{region 'Documentation'}
(*!
<summary>Calls Preparations and supplies their scenario-specific combined observations.</summary>
<description>
Called after ProcessAbort on every initialized call except Completed, with the current
Preparation-phase Enable. Call Preparations even when disabled so their observations and
deactivation remain correct; report the combination through UpdatePreparationStatus.

Only enabled phase processing may advance through NextPreparationState or
CompletePreparations. After entry into Test states, loss of Preparation Ready or Completed is not by
itself a Test Case failure. This abstract hook has no base implementation.
</description>
*)
{endregion}
METHOD PROTECTED ABSTRACT ProcessPreparations
VAR_INPUT
    Enable: BOOL; //! TRUE while this hook's lifecycle phase is active; FALSE must not advance that phase.
END_VAR
(* Example: declare a local ObservedStatus : ST_PreparationStatus; combine multiple Preparations as needed.
MyPreparation(Enable := Enable);
ObservedStatus := MyPreparation.Status;
UpdatePreparationStatus(Ready := ObservedStatus.Ready,
    Running := ObservedStatus.Running,
    Completed := ObservedStatus.Completed,
    HasError := ObservedStatus.Error,
    State := ObservedStatus.State);
IF Enable AND FPreparationStatus.Completed AND NOT FPreparationStatus.Error THEN
    CompletePreparations();
END_IF;
*)
END_METHOD

{region 'Documentation'}
(*!
<summary>Consumes same-task requests, reports each received request and prioritizes Reset &gt; Abort &gt; Start.</summary>
<description>
Discards requests before initialization; never changes lifecycle state.
</description>
*)
{endregion}
METHOD PRIVATE ProcessRequests
VAR_IN_OUT
    InputRequests : ST_Command; //! Same-task request mailbox consumed and cleared, including calls made before successful initialization.
END_VAR
VAR_OUTPUT
    Requests : ST_Command; //! Qualified request snapshot with Reset over Abort over Start; all FALSE before initialization.
END_VAR
Requests.Reset := FALSE;
Requests.Abort := FALSE;
Requests.Start := FALSE;

IF NOT FInitialized THEN
    InputRequests.Reset := FALSE;
    InputRequests.Abort := FALSE;
    InputRequests.Start := FALSE;
    RETURN;
END_IF;

Requests.Reset := InputRequests.Reset;
Requests.Abort := InputRequests.Abort AND NOT InputRequests.Reset;
Requests.Start := InputRequests.Start AND NOT InputRequests.Abort AND NOT InputRequests.Reset;

IF InputRequests.Reset THEN
    PublishEvent(Event := CreateResetEvent(OwnerScope := E_OwnerScope.TestCase,
        Name := FName,
        ResourceName := FResourceName,
        State := FState));
END_IF;

IF InputRequests.Abort THEN
    PublishEvent(Event := CreateAbortEvent(OwnerScope := E_OwnerScope.TestCase,
        Name := FName,
        ResourceName := FResourceName,
        State := FState));
END_IF;

IF InputRequests.Start THEN
    PublishEvent(Event := CreateStartEvent(OwnerScope := E_OwnerScope.TestCase,
        Name := FName,
        ResourceName := FResourceName,
        State := FState));
END_IF;

InputRequests.Reset := FALSE;
InputRequests.Abort := FALSE;
InputRequests.Start := FALSE;
END_METHOD

{region 'Documentation'}
(*!
<summary>Resets owned scenario resources and Assertions during the Reset phase.</summary>
<description>
Called after the base restores the Preparation snapshot to Unknown. Request Assertion resets;
their next regular calls process those requests with bound inputs. Finish through CompleteReset only
once the owned reset work is complete.

Preserve configuration and publisher bindings. One-shot resource protocols must not be
retriggered every cycle. The base owns ResetTimeout; this abstract hook has no base
implementation.
</description>
*)
{endregion}
METHOD PROTECTED ABSTRACT ProcessReset
(* Example: request child resets and observe completion without blocking.
MyAssertion.Reset();
IF OwnedResourcesReset THEN
    CompleteReset();
END_IF;
Issue one-shot resource requests only once if their protocol requires it.
*)
END_METHOD

{region 'Documentation'}
(*!
<summary>Performs scenario actions in the current Test state.</summary>
<description>
Called after ProcessPreparations on every initialized call except Completed. Enable reflects
the phase at invocation, including transitions made by earlier hooks. Keep required cyclic resource
calls active while disabled, but do not advance the Test phase.

Use NextTestState and CompleteTests for immediate transitions. Check errors before successful
completion; do not rely on a previously cached phase flag after changing state. This abstract hook
has no base implementation.
</description>
*)
{endregion}
METHOD PROTECTED ABSTRACT ProcessTests
VAR_INPUT
    Enable: BOOL; //! TRUE while this hook's lifecycle phase is active; FALSE must not advance that phase.
END_VAR
(* Example: keep required cyclic object calls outside the Enable guard.
MyTestObject();
IF NOT Enable THEN
    RETURN;
END_IF;
Perform the action for the current State; check errors before completion.
IF TestCompleted THEN
    CompleteTests();
END_IF;
*)
END_METHOD

{region 'Documentation'}
(*!
<summary>Publishes through the selected instance publisher; the buffer owns lost-event accounting.</summary>
*)
{endregion}
METHOD PRIVATE PublishEvent
VAR_INPUT
    Event : ST_Event; //! Payload copied once through the selected usable publisher, which assigns sequence/time and accounts for loss.
END_VAR
EventPublisher.PublishEvent(Event := Event);
END_METHOD

{region 'Documentation'}
(*!
<summary>Records an Abort request for the next regular FB call.</summary>
<description>
Repeated positive calls coalesce in the same-task request storage. Processing consumes the
requests with priority Reset, Abort, Start; calls before successful initialization are discarded
when processed.

Abort requests controlled termination of execution, not Reset cancellation. The owner
lifecycle determines whether the request applies.
</description>
*)
{endregion}
METHOD PUBLIC RequestAbort
FMethodRequests.Abort := TRUE;
END_METHOD

{region 'Documentation'}
(*!
<summary>Records a Reset request for the next regular FB call.</summary>
<description>
Repeated positive calls coalesce in the same-task request storage. Processing consumes the
requests with priority Reset, Abort, Start; calls before successful initialization are discarded
when processed.

Lifecycle Reset preserves configuration and publisher binding. It is not reinitialization or
Event Buffer Reset; capacity admission belongs to the parent when this object is a child.
</description>
*)
{endregion}
METHOD PUBLIC RequestReset
FMethodRequests.Reset := TRUE;
END_METHOD

{region 'Documentation'}
(*!
<summary>Records a Start request for the next regular FB call.</summary>
<description>
Repeated positive calls coalesce in the same-task request storage. Processing consumes the
requests with priority Reset, Abort, Start; calls before successful initialization are discarded
when processed.

Start is accepted by the lifecycle only in ready Idle. Recording the request does not start
execution synchronously.
</description>
*)
{endregion}
METHOD PUBLIC RequestStart
FMethodRequests.Start := TRUE;
END_METHOD

{region 'Documentation'}
(*!
<summary>Own contribution to the global Event Buffer reservation; changed only with that
aggregate.</summary>
*)
{endregion}
{attribute 'monitoring' := 'call'}
PROPERTY PUBLIC ReservedEntryCount : UINT //! Own contribution to the global Event Buffer reservation; changed only with that aggregate.
GET // PUBLIC
ReservedEntryCount := FReservedEntryCount;
END_GET
END_PROPERTY

{region 'Documentation'}
(*!
<summary>Adjusts this owner's reservation to its execution budget immediately.</summary>
<description>
The budget uses configured state counts and the collected AssertionCountTotal, which must be
valid and stable before Start. Local contribution and publisher accounting are updated together
without a lifecycle transition.

Accepted permits dispatch; WaitingForCapacity is retryable under the owner's timeout; Error
denotes invalid setup or an impossible budget. Calling before initialization reports a Framework
error. Repeated success aligns the total rather than adding a second budget.
</description>
*)
{endregion}
METHOD PUBLIC FINAL ReserveExecutionEvents : E_EventReservationResult //! Accepted on success, WaitingForCapacity for retryable pressure, Error for invalid setup or an impossible budget.
VAR
    EntryCount : UDINT;
END_VAR
VAR CONSTANT
    FixedEventCount : UDINT := 9;
    MaxReservationEntryCount : UDINT := 65535;
END_VAR
ReserveExecutionEvents := E_EventReservationResult.Error;
IF NOT FInitialized THEN
    PublishEvent(Event := CreateFrameworkEvent(Name := FName,
        ResourceName := FResourceName,
        State := FState,
        Severity := E_EventSeverity.Error,
        Message := 'ReserveExecutionEvents requires an initialized Test Case.'));
    RETURN;
END_IF;

EntryCount := INT_TO_UDINT(FPreparationStateCount)
    + INT_TO_UDINT(FTestStateCount)
    + UINT_TO_UDINT(FStatus.AssertionCountTotal)
    + FixedEventCount;
IF EntryCount > MaxReservationEntryCount THEN
    PublishEvent(Event := CreateFrameworkEvent(Name := FName,
        ResourceName := FResourceName,
        State := FState,
        Severity := E_EventSeverity.Error,
        Message := 'Test Case event budget exceeds the reservation range.'));
    RETURN;
END_IF;

ReserveExecutionEvents := UpdateEventReservation(EntryCount := UDINT_TO_UINT(EntryCount),
    HeadroomEntryCount := Param_EventBuffer.EventBufferExecutionHeadroom,
    ConcurrentEntryCount := GVL_Constants.TestSuiteExecutionEventCount);
END_METHOD

{region 'Documentation'}
(*!
<summary>Adjusts this owner's reservation for capacity-admitted Reset immediately.</summary>
<description>
Does not dispatch Reset or clear existing events. Shared headroom and the Suite allowance
participate in admission, not this owner's stored contribution.

Accepted, WaitingForCapacity and Error distinguish success, temporary pressure and invalid
setup. An uninitialized call reports a Framework error. Lifecycle Reset must not silently clear the
reservation.
</description>
*)
{endregion}
METHOD PUBLIC FINAL ReserveResetEvents : E_EventReservationResult //! Accepted on success, WaitingForCapacity for retryable pressure, Error for invalid setup or an impossible budget.
ReserveResetEvents := E_EventReservationResult.Error;
IF NOT FInitialized THEN
    PublishEvent(Event := CreateFrameworkEvent(Name := FName,
        ResourceName := FResourceName,
        State := FState,
        Severity := E_EventSeverity.Error,
        Message := 'ReserveResetEvents requires an initialized Test Case.'));
    RETURN;
END_IF;

ReserveResetEvents := UpdateEventReservation(EntryCount := GVL_Constants.TestCaseResetEventCount,
    HeadroomEntryCount := Param_EventBuffer.EventBufferResetHeadroom,
    ConcurrentEntryCount := GVL_Constants.TestSuiteResetEventCount);
END_METHOD

{region 'Documentation'}
(*!
<summary>Current held Test Case result.</summary>
*)
{endregion}
{attribute 'monitoring' := 'call'}
PROPERTY PUBLIC Result : E_Result //! Current held Test Case result.
GET // PUBLIC
Result := FResult;
END_GET
END_PROPERTY

{region 'Documentation'}
(*!
<summary>Selects lifecycle transitions from requests, observations and timeout supervision.</summary>
*)
{endregion}
METHOD PRIVATE Sequencer
VAR_INPUT
    Requests : ST_Command; //! Consumed request snapshot whose applicability is evaluated against current lifecycle state and error/timeout priority.
END_VAR
VAR
    Message : STRING(GVL_Constants.MessageLength);
END_VAR
IF NOT FInitialized THEN
    IF FState <> E_State.Uninitialized THEN
        ChangeState(NewState := E_State.Uninitialized);
    END_IF;
    RETURN;
END_IF;
IF Requests.Reset THEN
    ChangeState(NewState := E_State.Reset);
END_IF;

CASE FState OF
    E_State.Uninitialized:
        RETURN;

    E_State.Reset:
        IF NOT FStateTimer.IsValid THEN
            PublishEvent(Event := CreateFrameworkEvent(Name := FName,
                ResourceName := FResourceName,
                State := FState,
                Severity := E_EventSeverity.Error,
                Message := 'Task clock error during Test Case reset.'));
            FResult := E_Result.Error;
            ChangeState(NewState := E_State.Completing);
            RETURN;
        END_IF;
        IF FStateTimer.ElapsedLTime >= TIME_TO_LTIME(FConfig.ResetTimeout) THEN
            FHasResetTimeout := TRUE;
            PublishEvent(Event := CreateFrameworkEvent(Name := FName,
                ResourceName := FResourceName,
                State := FState,
                Severity := E_EventSeverity.Error,
                Message := 'Test Case reset timeout reached.'));
            FResult := E_Result.Error;
            ChangeState(NewState := E_State.Completing);
            RETURN;
        END_IF;
        RETURN;

    E_State.Idle:
        IF Requests.Start AND NOT Requests.Abort AND IsReady THEN
            ChangeState(NewState := E_State.Starting);
        END_IF;
        RETURN;

    E_State.Starting:
        IF FResult = E_Result.Error THEN
            ChangeState(NewState := E_State.AbortingFromError);
            RETURN;
        END_IF;
        IF FPreparationStatus.Error THEN
            Message := CONCAT('Preparation error. Preparation state = ', INT_TO_STRING(FPreparationStatus.State));
            Error(Message := Message);
            RETURN;
        END_IF;
        IF FAggregator.Result = E_Result.Error THEN
            Error(Message := 'Test Case evaluation reported Error.');
            RETURN;
        END_IF;
        IF NOT FExecutionTimer.IsValid OR NOT FStateTimer.IsValid THEN
            Error(Message := 'Task clock error.');
            RETURN;
        END_IF;
        IF FExecutionTimer.ElapsedLTime >= TIME_TO_LTIME(FConfig.Timeout) THEN
            FHasTimeout := TRUE;
            Error(Message := 'Test Case timeout.');
            RETURN;
        END_IF;
        IF Requests.Abort THEN
            ChangeState(NewState := E_State.Aborting);
            RETURN;
        END_IF;
        IF (FPreparationStateCount = 0) OR FPreparationStatus.Completed THEN
            ChangeState(NewState := E_State.Running);
            RETURN;
        END_IF;
        ChangeState(NewState := E_State.Preparing);
        RETURN;

    E_State.Preparing..(E_State.Running - 1):
        IF FResult = E_Result.Error THEN
            ChangeState(NewState := E_State.AbortingFromError);
            RETURN;
        END_IF;
        IF NOT IsPreparationActive THEN
            Message := CONCAT('Invalid preparation state = ', INT_TO_STRING(FState));
            Error(Message := Message);
            RETURN;
        END_IF;
        IF FPreparationStatus.Error THEN
            Message := CONCAT('Preparation error. Preparation state = ', INT_TO_STRING(FPreparationStatus.State));
            Error(Message := Message);
            RETURN;
        END_IF;
        IF FAggregator.Result = E_Result.Error THEN
            Error(Message := 'Test Case evaluation reported Error.');
            RETURN;
        END_IF;
        IF NOT FExecutionTimer.IsValid OR NOT FStateTimer.IsValid THEN
            Error(Message := 'Task clock error.');
            RETURN;
        END_IF;
        IF FStateTimer.ElapsedLTime >= TIME_TO_LTIME(FConfig.PreparationTimeout) THEN
            FHasPreparationTimeout := TRUE;
            Message := CONCAT('Preparation timeout. Preparation state = ', INT_TO_STRING(FPreparationStatus.State));
            Error(Message := Message);
            RETURN;
        END_IF;
        IF FExecutionTimer.ElapsedLTime >= TIME_TO_LTIME(FConfig.Timeout) THEN
            FHasTimeout := TRUE;
            Error(Message := 'Test Case timeout.');
            RETURN;
        END_IF;
        IF Requests.Abort THEN
            ChangeState(NewState := E_State.Aborting);
            RETURN;
        END_IF;
        IF (FPreparationStateCount = 0) OR FPreparationStatus.Completed THEN
            ChangeState(NewState := E_State.Running);
            RETURN;
        END_IF;
        // Leave to Running by CompletePreparations
        RETURN;

    E_State.Running..(E_State.Completing - 1):
        IF FResult = E_Result.Error THEN
            ChangeState(NewState := E_State.AbortingFromError);
            RETURN;
        END_IF;
        IF NOT IsTestingActive THEN
            Message := CONCAT('Invalid testing state = ', INT_TO_STRING(FState));
            Error(Message := Message);
            RETURN;
        END_IF;
        IF FAggregator.Result = E_Result.Error THEN
            Error(Message := 'Test Case evaluation reported Error.');
            RETURN;
        END_IF;
        IF NOT FExecutionTimer.IsValid THEN
            Error(Message := 'Task clock error.');
            RETURN;
        END_IF;
        IF FExecutionTimer.ElapsedLTime >= TIME_TO_LTIME(FConfig.Timeout) THEN
            FHasTimeout := TRUE;
            Error(Message := 'Test Case timeout.');
            RETURN;
        END_IF;
        IF Requests.Abort THEN
            ChangeState(NewState := E_State.Aborting);
            RETURN;
        END_IF;
        // Leave to Completing by CompleteTests
        RETURN;

    E_State.Completing:
        ChangeState(NewState := E_State.Completed);
        RETURN;

    E_State.Completed:
        // Leave to Reset on ResetRequested.
        RETURN;

    E_State.Aborting, E_State.AbortingFromError:
        IF NOT FStateTimer.IsValid THEN
            PublishEvent(Event := CreateFrameworkEvent(Name := FName,
                ResourceName := FResourceName,
                State := FState,
                Severity := E_EventSeverity.Error,
                Message := 'Task clock error during Test Case abort.'));
            FResult := E_Result.Error;
            ChangeState(NewState := E_State.Completing);
            RETURN;
        END_IF;
        IF FStateTimer.ElapsedLTime >= TIME_TO_LTIME(FConfig.AbortTimeout) THEN
            FHasAbortTimeout := TRUE;
            PublishEvent(Event := CreateFrameworkEvent(Name := FName,
                ResourceName := FResourceName,
                State := FState,
                Severity := E_EventSeverity.Error,
                Message := 'Test Case abort timeout reached.'));
            FResult := E_Result.Error;
            ChangeState(NewState := E_State.Completing);
            RETURN;
        END_IF;
        IF (FState = E_State.Aborting) AND (FResult = E_Result.Error) THEN
            ChangeState(NewState := E_State.AbortingFromError);
        END_IF;
        RETURN;

    E_State.Aborted, E_State.Error:
        Error(Message := 'Unexpected legacy lifecycle state.');
        RETURN;
ELSE
    Error(Message := 'Unhandled Test Case lifecycle state.');
END_CASE;
END_METHOD

{region 'Documentation'}
(*!
<summary>Current Test Case lifecycle state.</summary>
*)
{endregion}
{attribute 'monitoring' := 'call'}
PROPERTY PUBLIC State : E_State //! Current Test Case lifecycle state.
GET // PUBLIC
State := FState;
END_GET
END_PROPERTY

{region 'Documentation'}
(*!
<summary>Returns the latest Test Case status snapshot without executing children.</summary>
<description>
The base refreshes this snapshot on every FB call, including Uninitialized and Completed.
Assertion counters come from the current collection; the completed owner result remains held.
Runtime is TIME.

Preparation observations are available separately through PreparationStatus. Optional external
publication requires an explicit data wrapper, not access to owner instance data.
</description>
*)
{endregion}
PROPERTY PUBLIC Status : ST_TestCaseStatus //! Returns the latest Test Case status snapshot without executing children.
GET // PUBLIC
Status := FStatus;
END_GET
END_PROPERTY

{region 'Documentation'}
(*!
<summary>Reports the configured maximum number of Test-state entries along one finite lifecycle
path.</summary>
<description>
Set the backing field explicitly in Configure. Before configuration it is
StateCountNotConfigured (-1). Branches use the longest path, including bounded repeated entries;
this is not a count of child instances. Keep it fixed through execution.

At least one Test state is required. CheckInitialization bounds the value by
E_State.Completing - E_State.Running.
</description>
*)
{endregion}
{attribute 'monitoring' := 'call'}
PROPERTY PUBLIC TestStateCount : INT //! Reports the configured maximum number of Test-state entries along one finite lifecycle path.
GET // PUBLIC
TestStateCount := FTestStateCount;
END_GET
END_PROPERTY

{region 'Documentation'}
(*!
<summary>Checks target capacity before changing either reservation count; zero releases without capacity gating.</summary>
<description>
A zero target with no existing contribution succeeds without accessing a publisher. Releasing a nonzero contribution delegates to FreeReservedSpace without a free-capacity check. Positive targets first require valid publisher/accounting and permanent capacity for target plus the concurrent Suite allowance plus headroom. Temporary free capacity uses aggregate minus old own contribution plus target plus headroom; it does not add the Suite allowance again. Even unchanged or reduced positive targets must pass those checks. Failure leaves both ledgers unchanged.
</description>
*)
{endregion}
METHOD PRIVATE UpdateEventReservation : E_EventReservationResult //! Accepted after aligning the own contribution, WaitingForCapacity for temporary pressure, Error for invalid binding/accounting or impossible capacity.
VAR_INPUT
    EntryCount : UINT; //! Target total own reservation, not an additional delta; zero releases the complete own contribution.
    HeadroomEntryCount : UINT; //! Shared unreserved producer headroom included in permanent and temporary capacity checks for a nonzero target.
    ConcurrentEntryCount : UINT; //! Suite allowance used only in the permanent capacity check; actual temporary reservations already include the parent's contribution.
END_VAR
VAR
    Publisher : I_EventPublisher;
    RequiredCapacity : UDINT;
    RequiredFreeEntries : UDINT;
END_VAR
UpdateEventReservation := E_EventReservationResult.Error;
IF (EntryCount = 0) AND (FReservedEntryCount = 0) THEN
    UpdateEventReservation := E_EventReservationResult.Accepted;
    RETURN;
END_IF;

Publisher := EventPublisher;

IF EntryCount = 0 THEN
    IF Publisher.FreeReservedSpace(EntryCount := FReservedEntryCount,
        OwnerReservedEntryCount := FReservedEntryCount) THEN
        UpdateEventReservation := E_EventReservationResult.Accepted;
    END_IF;
    RETURN;
END_IF;

IF NOT Publisher.IsValid THEN
    RETURN;
END_IF;
RequiredCapacity := UINT_TO_UDINT(EntryCount)
    + UINT_TO_UDINT(ConcurrentEntryCount)
    + UINT_TO_UDINT(HeadroomEntryCount);
IF RequiredCapacity > UINT_TO_UDINT(Publisher.Capacity) THEN
    RETURN;
END_IF;
IF FReservedEntryCount > Publisher.ReservedEntryCount THEN
    RETURN;
END_IF;

RequiredFreeEntries := UINT_TO_UDINT(Publisher.ReservedEntryCount)
    - UINT_TO_UDINT(FReservedEntryCount)
    + UINT_TO_UDINT(EntryCount)
    + UINT_TO_UDINT(HeadroomEntryCount);
IF RequiredFreeEntries > UINT_TO_UDINT(Publisher.FreeEntryCount) THEN
    UpdateEventReservation := E_EventReservationResult.WaitingForCapacity;
    RETURN;
END_IF;

IF EntryCount < FReservedEntryCount THEN
    IF Publisher.FreeReservedSpace(EntryCount := FReservedEntryCount - EntryCount,
        OwnerReservedEntryCount := FReservedEntryCount) THEN
        UpdateEventReservation := E_EventReservationResult.Accepted;
    END_IF;
    RETURN;
END_IF;

IF Publisher.ReserveSpace(EntryCount := EntryCount - FReservedEntryCount,
    HeadroomEntryCount := HeadroomEntryCount,
    OwnerReservedEntryCount := FReservedEntryCount) THEN
    UpdateEventReservation := E_EventReservationResult.Accepted;
ELSE
    UpdateEventReservation := E_EventReservationResult.WaitingForCapacity;
END_IF;
END_METHOD

{region 'Documentation'}
(*!
<summary>Replaces the combined Preparation observations without calling children.</summary>
<description>
Combine multiple Preparations according to the concrete scenario; this method imposes no
universal AND/OR aggregation. All supplied flags replace previous observations; Ready is suppressed
while Running.

ExecutionStatus follows Error, Completed, Running, then Idle when Ready and NotReady
otherwise. State is optional diagnostic context, not the owner's phase. Initial/reset Unknown
snapshots are established separately by the base.
</description>
*)
{endregion}
METHOD PROTECTED UpdatePreparationStatus
VAR_INPUT
    Ready : BOOL; //! Resource can be driven to the target state; suppressed while Running. Does not mean target reached.
    Running : BOOL; //! Preparation is actively driving the resource toward its target; forces Ready to FALSE.
    Completed : BOOL; //! Preparation target is currently reached; observation is not latched.
    HasError : BOOL; //! Preparation cannot continue meaningfully; reported as an error observation.
    State : E_State := E_State.Uninitialized; //! Optional combined Preparation state for observation; default Uninitialized.
END_VAR
FPreparationStatus.State := State;
FPreparationStatus.Ready := Ready AND NOT Running;
FPreparationStatus.Running := Running;
FPreparationStatus.Completed := Completed;
FPreparationStatus.Error := HasError;

IF HasError THEN
    FPreparationStatus.ExecutionStatus := E_ExecutionStatus.Error;
ELSIF Completed THEN
    FPreparationStatus.ExecutionStatus := E_ExecutionStatus.Completed;
ELSIF Running THEN
    FPreparationStatus.ExecutionStatus := E_ExecutionStatus.Running;
ELSIF Ready THEN
    FPreparationStatus.ExecutionStatus := E_ExecutionStatus.Idle;
ELSE
    FPreparationStatus.ExecutionStatus := E_ExecutionStatus.NotReady;
END_IF;
END_METHOD

{region 'Documentation'}
(*!
<summary>Applies lifecycle-specific owner result rules to the current aggregate.</summary>
*)
{endregion}
METHOD PRIVATE UpdateResult
IF (FResult = E_Result.Error) AND (FState <> E_State.Uninitialized) THEN
    RETURN;
END_IF;

CASE FState OF
    E_State.Uninitialized, E_State.Starting:
        FResult := E_Result.NotEvaluated;
    E_State.Reset, E_State.Idle:
        RETURN;
    E_State.Aborting:
        IF (FResult = E_Result.Error) OR (FAggregator.Result = E_Result.Error) THEN
            FResult := E_Result.Error;
        ELSE
            FResult := E_Result.Abort;
        END_IF;
    E_State.AbortingFromError:
        FResult := E_Result.Error;
    E_State.Completing:
        IF (FResult = E_Result.Error) OR (FAggregator.Result = E_Result.Error) THEN
            FResult := E_Result.Error;
            RETURN;
        END_IF;
        IF FResult = E_Result.Abort THEN
            RETURN;
        END_IF;
        CASE FAggregator.Result OF
            E_Result.Failed:
                FResult := E_Result.Failed;
            E_Result.Passed, E_Result.NotEvaluated:
                FResult := E_Result.Passed;
        ELSE
            FResult := E_Result.Error;
        END_CASE;
    E_State.Completed:
        RETURN;
ELSE
    IF IsPreparationActive OR IsTestingActive THEN
        FResult := E_Result.NotEvaluated;
    ELSE
        FResult := E_Result.Error;
    END_IF;
END_CASE;
END_METHOD

{region 'Documentation'}
(*!
<summary>Refreshes the typed snapshot from current lifecycle state; does not invoke children.</summary>
*)
{endregion}
METHOD PRIVATE UpdateStatus
VAR
    ExecutionStatus : ST_TestCaseExecutionStatus;
END_VAR
ExecutionStatus.State := FState;
ExecutionStatus.Result := FResult;
ExecutionStatus.ConfigError := FConfigError;
CASE FState OF
    E_State.Uninitialized:
        ExecutionStatus.ExecutionStatus := E_ExecutionStatus.NotReady;
        ExecutionStatus.Uninitialized := TRUE;
    E_State.Reset:
        ExecutionStatus.ExecutionStatus := E_ExecutionStatus.Reset;
    E_State.Idle:
        ExecutionStatus.ExecutionStatus := E_ExecutionStatus.Idle;
        ExecutionStatus.Ready := IsReady;
    E_State.Starting:
        ExecutionStatus.ExecutionStatus := E_ExecutionStatus.Starting;
    E_State.Completing:
        ExecutionStatus.ExecutionStatus := E_ExecutionStatus.Completing;
    E_State.Completed:
        ExecutionStatus.ExecutionStatus := E_ExecutionStatus.Completed;
        ExecutionStatus.Completed := TRUE;
        ExecutionStatus.Aborted := FResult = E_Result.Abort;
        ExecutionStatus.Error := FResult = E_Result.Error;
    E_State.Aborting, E_State.AbortingFromError:
        ExecutionStatus.ExecutionStatus := E_ExecutionStatus.Aborting;
ELSE
    IF IsPreparationActive OR IsTestingActive THEN
        ExecutionStatus.ExecutionStatus := E_ExecutionStatus.Running;
        ExecutionStatus.Running := TRUE;
        ExecutionStatus.PreparationActive := IsPreparationActive;
        ExecutionStatus.TestActive := IsTestingActive;
    ELSE
        ExecutionStatus.ExecutionStatus := E_ExecutionStatus.Error;
        ExecutionStatus.Error := TRUE;
    END_IF;
END_CASE;
ExecutionStatus.Error := HasError;
FStatus.Execution := ExecutionStatus;
FStatus.PreparationStateCount := 0;
IF (FPreparationStateCount >= 0)
    AND (FPreparationStateCount <= E_State.Running - E_State.Preparing) THEN
    FStatus.PreparationStateCount := INT_TO_UINT(FPreparationStateCount);
END_IF;
FStatus.TestStateCount := 0;
IF (FTestStateCount >= 1)
    AND (FTestStateCount <= E_State.Completing - E_State.Running) THEN
    FStatus.TestStateCount := INT_TO_UINT(FTestStateCount);
END_IF;
FStatus.Runtime := FExecutionTimer.ElapsedTime;
FStatus.AssertionCountTotal := FAggregator.TotalCount;
FStatus.AssertionCountPassed := FAggregator.PassedCount;
FStatus.AssertionCountFailed := FAggregator.FailedCount;
FStatus.AssertionCountError := FAggregator.ErrorCount;
END_METHOD

END_FUNCTION_BLOCK

// ---- Framework/EventBuffer/POU/AggregationEvents/CreateTestCaseAggregationEvent.TcPOU
{region 'Documentation'}
(*!
<summary>Constructs a Test Case aggregation event from an already aggregated status snapshot.</summary>
<description>
Runtime is rendered as unsigned milliseconds; the caller owns publication.


Compact JSON fields are total, passed, failed, error and runtime. Counts and runtime are unsigned decimal numbers. This formats the supplied snapshot without validating completion or recomputing aggregation; the owner controls finalization order and publication.
</description>
*)
{endregion}
FUNCTION CreateTestCaseAggregationEvent : ST_Event //! Constructed event value; not published. The publisher assigns SequenceId and Timestamp.
VAR_INPUT
    Name : STRING(GVL_Constants.NameLength); //! Hierarchical owner name used to identify events; must satisfy the naming contract.
    ResourceName : STRING(GVL_Constants.ResourceNameLength) := ''; //! Optional resource context for diagnostics; empty by default.
    Status : ST_TestCaseStatus; //! Already aggregated owner status snapshot; the function formats it without observing children.
END_VAR
VAR
    RuntimeMilliseconds : UDINT;
END_VAR

RuntimeMilliseconds := TIME_TO_UDINT(Status.Runtime);

CreateTestCaseAggregationEvent.SequenceId := 0;
CreateTestCaseAggregationEvent.Timestamp := 0;
CreateTestCaseAggregationEvent.OwnerScope := E_OwnerScope.TestCase;
CreateTestCaseAggregationEvent.EventType := E_EventType.Aggregation;
CreateTestCaseAggregationEvent.Severity := SelectResultSeverity(Result := Status.Execution.Result);
CreateTestCaseAggregationEvent.Name := Name;
CreateTestCaseAggregationEvent.ResourceName := ResourceName;
CreateTestCaseAggregationEvent.State := Status.Execution.State;
CreateTestCaseAggregationEvent.Result := Status.Execution.Result;

CreateTestCaseAggregationEvent.Message := CONCAT(STR1 := '{"total":',
    STR2 := UINT_TO_STRING(Status.AssertionCountTotal));
CreateTestCaseAggregationEvent.Message := CONCAT(STR1 := CreateTestCaseAggregationEvent.Message,
    STR2 := ',"passed":');
CreateTestCaseAggregationEvent.Message := CONCAT(STR1 := CreateTestCaseAggregationEvent.Message,
    STR2 := UINT_TO_STRING(Status.AssertionCountPassed));
CreateTestCaseAggregationEvent.Message := CONCAT(STR1 := CreateTestCaseAggregationEvent.Message,
    STR2 := ',"failed":');
CreateTestCaseAggregationEvent.Message := CONCAT(STR1 := CreateTestCaseAggregationEvent.Message,
    STR2 := UINT_TO_STRING(Status.AssertionCountFailed));
CreateTestCaseAggregationEvent.Message := CONCAT(STR1 := CreateTestCaseAggregationEvent.Message,
    STR2 := ',"error":');
CreateTestCaseAggregationEvent.Message := CONCAT(STR1 := CreateTestCaseAggregationEvent.Message,
    STR2 := UINT_TO_STRING(Status.AssertionCountError));
CreateTestCaseAggregationEvent.Message := CONCAT(STR1 := CreateTestCaseAggregationEvent.Message,
    STR2 := ',"runtime":');
CreateTestCaseAggregationEvent.Message := CONCAT(STR1 := CreateTestCaseAggregationEvent.Message,
    STR2 := UDINT_TO_STRING(RuntimeMilliseconds));
CreateTestCaseAggregationEvent.Message := CONCAT(STR1 := CreateTestCaseAggregationEvent.Message, STR2 := '}');

END_FUNCTION

// ---- Framework/Assertions/POU/BasicTypes/Bool/AssertTrue.TcPOU
{region 'Documentation'}
(*!
<summary>Checks that the BOOL value is TRUE.</summary>
*)
{endregion}
FUNCTION_BLOCK AssertTrue EXTENDS AssertionBase
VAR_INPUT
    IN : BOOL; //! Actual value checked or observed by this Assertion.
END_VAR

SUPER^();

{region 'Documentation'}
(*!
<summary>Evaluate whether the BOOL value is TRUE.</summary>
*)
{endregion}
METHOD PROTECTED Assert
VAR
    Message : STRING(GVL_Constants.MessageLength);
    ActualText : STRING(GVL_Constants.AssertionValueLength);
END_VAR
IF NOT EvaluationActive THEN
    RETURN;
END_IF;

IF Result = E_Result.Error THEN
    RETURN;
END_IF;

IF Result = E_Result.Failed THEN
    RETURN;
END_IF;

IF NOT IN THEN
    ActualText := BOOL_TO_STRING(IN);
    Message := CONCAT('Assertion failed: values are not equal. Expected = TRUE, Actual = ',
        ActualText);
    Message := CONCAT(Message, '.');
    Fail(Message := Message);
    RETURN;
END_IF;

Pass();
END_METHOD

END_FUNCTION_BLOCK

// ---- Framework/Assertions/POU/AssertionBase.TcPOU
{region 'Documentation'}
(*!
<summary>Shared cyclic assertion lifecycle, identity and monotonic result escalation.</summary>
<description>

Initialize from the owning Test Case configuration, then call the concrete FB once per
cycle with its typed inputs. Derived FB bodies call SUPER^() once. The base invokes Assert only
after successful initialization and outside a reset call.

Enable controls observation. ObserveFirstCycle determines whether its first enabled call
is observed. EvaluationActive normally follows ObservationActive; explicit-evaluation and
history-based families refine this gate.

Reset queues work for the next FB call: result becomes NotEvaluated, observation history
is cleared by ResetAssertion and that call performs no assertion check. Identity and publisher
binding are retained. Initialize also queues this reset, including when initialization
fails.

Pass cannot clear Failed or Error. Fail escalates NotEvaluated or Passed; Error can also
escalate Failed. Findings are published once per result escalation, not every cyclic failure. A
failed publication is not retried.

State is owner-supplied finding context, not a state machine input. Diagnostic value text
may be shortened or rounded; comparisons use the original typed values. The selected publisher
must exist before any publication.

</description>
*)
{endregion}
FUNCTION_BLOCK ABSTRACT AssertionBase IMPLEMENTS I_Assertion
VAR_INPUT
    Enable : BOOL; //! Enables observation; Initialize's ObserveFirstCycle setting controls the first enabled call.
    State : E_State := E_State.Uninitialized; //! Owner's current lifecycle state included in finding events; default Uninitialized.
END_VAR
VAR
    /// Instance binding selected by BindPublisher or lazily by EventPublisher.
    FEventPublisher : I_EventPublisher;
    FName : STRING(GVL_Constants.NameLength) := '<UnnamedAssertion>';
    FResourceName : STRING(GVL_Constants.ResourceNameLength);
    FResult : E_Result := E_Result.NotEvaluated;
    FEnabled : BOOL;
    FInitialized : BOOL;
    FResetRequested : BOOL;
    FObserveFirstCycle : BOOL := TRUE;
    FEnablePrevious : BOOL;
    FResetActive : BOOL;
END_VAR

FEnablePrevious := FEnabled AND NOT FResetActive;
FEnabled := Enable;
FResetActive := FResetRequested;

IF FResetActive THEN
    FResetRequested := FALSE;
    FEnablePrevious := FALSE;
    FResult := E_Result.NotEvaluated;
    ResetAssertion();
    RETURN;
END_IF;

IF NOT FInitialized THEN
    RETURN;
END_IF;

Assert();

{region 'Documentation'}
(*!
<summary>Implement the typed observation and result check.</summary>
<description>

Called once per initialized non-reset FB call, including disabled calls. Apply the
family-specific ObservationActive and EvaluationActive gates. Validate prerequisites before
access; applicable Error checks precede Failed checks and Pass is the successful
fallback.

Do not suppress required observation or configuration-error checks merely because Result
is Failed. The implementation comment provides an illustrative ordering, not mandatory test
conditions.

</description>
*)
{endregion}
METHOD PROTECTED ABSTRACT Assert
(*
Implementation sketch, not a mandatory copy template.
Keep applicable Error checks before Failed checks; Pass is the fallback.
Omit conditions that do not exist. Multiple branches per severity are allowed.

Before result evaluation:
- Perform required observation/snapshot work under its own activity gate.
- Validate each operation's prerequisites before accessing its data.
- Observation errors may occur without EvaluationActive.
- Do not skip required observation or memory safety checks because of Result.
- Validate independent initialization/configuration when it is performed;
  do not report unused inputs as errors merely because the FB is called.

Example result evaluation (placeholder conditions/messages):

IF NOT EvaluationActive THEN
    RETURN;
END_IF;

IF Result = E_Result.Error THEN
    RETURN;
END_IF;

IF ErrorConditionA THEN
    Error(Message := ErrorMessageA);
    RETURN;
END_IF;

IF ErrorConditionB THEN
    Error(Message := ErrorMessageB);
    RETURN;
END_IF;

IF Result = E_Result.Failed THEN
    RETURN;
END_IF;

IF FailureConditionA THEN
    Fail(Message := FailureMessageA);
    RETURN;
END_IF;

IF FailureConditionB THEN
    Fail(Message := FailureMessageB);
    RETURN;
END_IF;

Pass();

A held Failed result must not bypass applicable Error checks.
Pass/Fail/Error retain the monotonic result and suppress repeated findings.
*)
END_METHOD

{region 'Documentation'}
(*!
<summary>Select the instance publisher immediately; ignore a zero assignment.</summary>
<description>

Retains identity, result and observation state. The caller owns the service lifetime.
There is no lifecycle guard, reset or replay when replacing this binding.

</description>
*)
{endregion}
METHOD PUBLIC BindPublisher
VAR_INPUT
    Publisher : I_EventPublisher; //! Publisher retained by the Assertion; caller owns its lifetime. Zero leaves the current binding unchanged.
END_VAR
IF Publisher = 0 THEN
    RETURN;
END_IF;

FEventPublisher := Publisher;
END_METHOD

{region 'Documentation'}
(*!
<summary>Enable accepted at the last FB call; not proof of evaluation.</summary>
*)
{endregion}
{attribute 'monitoring' := 'call'}
PROPERTY PUBLIC Enabled : BOOL //! Enable accepted at the last FB call; not proof of evaluation.
GET // PUBLIC
Enabled := FEnabled;
END_GET
END_PROPERTY

{region 'Documentation'}
(*!
<summary>Escalate any non-Error result to Error and publish one finding.</summary>
<description>

Failed can escalate to Error. Repeated Error calls do nothing. The result is stored
before publication; a publication failure is not retried.

</description>
*)
{endregion}
METHOD PROTECTED Error
VAR_INPUT
    Message : STRING(GVL_Constants.MessageLength); //! Diagnostic text for this finding; copied into the event within MessageLength.
END_VAR
VAR
    Finding : ST_Event;
    PublishResult : INT;
END_VAR
IF FResult = E_Result.Error THEN
    RETURN;
END_IF;

FResult := E_Result.Error;
Finding := CreateAssertionErrorEvent(Name := FName,
    ResourceName := FResourceName,
    State := State,
    Message := Message);
PublishResult := EventPublisher.PublishEvent(Event := Finding);
END_METHOD

{region 'Documentation'}
(*!
<summary>Use the polymorphic ObservationActive gate for direct result evaluation.</summary>
<description>

Explicit-evaluation and history-based descendants override this getter. A TRUE gate
permits checking; it does not mean the result is Passed or that this call has published a
finding.

</description>
*)
{endregion}
{attribute 'monitoring' := 'call'}
PROPERTY PUBLIC EvaluationActive : BOOL //! Effective gate for direct result evaluation; delegates to ObservationActive in this base.
GET // PUBLIC
EvaluationActive := ObservationActive;
END_GET
END_PROPERTY

{region 'Documentation'}
(*!
<summary>Return the instance publisher, binding the global default lazily if still
unset.</summary>
<description>

The first read without a local binding copies GVL_EventBuffer.Publisher. A nonzero local
binding is retained; later global changes do not replace it. This getter can therefore change
the binding. Publication requires a valid publisher.

</description>
*)
{endregion}
{attribute 'monitoring' := 'variable'}
PROPERTY PUBLIC EventPublisher : I_EventPublisher //! Instance publisher; the first unbound access adopts and retains the global default.
GET // PUBLIC
IF FEventPublisher = 0 THEN
    FEventPublisher := GVL_EventBuffer.Publisher;
END_IF;
EventPublisher := FEventPublisher;
END_GET
END_PROPERTY

{region 'Documentation'}
(*!
<summary>Escalate NotEvaluated or Passed to Failed and publish one finding.</summary>
<description>

Already Failed or Error is unchanged. The result is stored before publication; a
publication failure is not retried.

</description>
*)
{endregion}
METHOD PROTECTED Fail
VAR_INPUT
    Message : STRING(GVL_Constants.MessageLength); //! Diagnostic text for this finding; copied into the event within MessageLength.
END_VAR
VAR
    Finding : ST_Event;
    PublishResult : INT;
END_VAR
CASE FResult OF
    E_Result.NotEvaluated, E_Result.Passed:
        FResult := E_Result.Failed;
ELSE
    RETURN;
END_CASE;

Finding := CreateAssertionFailedEvent(Name := FName,
    ResourceName := FResourceName,
    State := State,
    Message := Message);
PublishResult := EventPublisher.PublishEvent(Event := Finding);
END_METHOD

{region 'Documentation'}
(*!
<summary>Configure the hierarchical identity and observation settings; return initialization
success.</summary>
<description>
The Parent Test Case identity must already be valid. The complete name consists of the
Parent's three hierarchy segments and a nonempty local Assertion suffix, which may contain
additional dots. It must fit NameLength; sibling uniqueness remains the caller's
responsibility. The parent interface is read here, not retained.
The composed name is length-limited into Name before validation of the unshortened name,
so an invalid name can remain available for diagnostics. Missing parent or invalid name
publishes a framework error and returns FALSE.
Clears base result and enable history and queues ResetAssertion for the next FB call,
where typed inputs are bound. ResourceName and ObserveFirstCycle are copied after a parent is
available. TRUE enables subsequent checking; normal Reset retains these settings.
</description>
*)
{endregion}
METHOD PUBLIC FINAL Initialize : BOOL //! TRUE after successful identity and setup validation; FALSE leaves the object uninitialized.
VAR_INPUT
    Parent : I_TestCase; //! Owning Test Case with an established Name; read during initialization, not retained.
    AssertionName : STRING(GVL_Constants.NameLength); //! Nonempty assertion suffix appended to Parent.Name; the complete name must satisfy the naming contract.
    ResourceName : STRING(GVL_Constants.ResourceNameLength) := ''; //! Optional resource context copied into finding events; empty by default.
    ObserveFirstCycle : BOOL := TRUE; //! TRUE observes the first enabled call; FALSE skips it. Default TRUE; does not delay explicit Evaluate.
END_VAR
VAR
    ParentName : STRING(GVL_Constants.NameLength);
    FullName : STRING(2 * GVL_Constants.NameLength + 1);
END_VAR
Initialize := FALSE;
FInitialized := FALSE;
FResult := E_Result.NotEvaluated;
FEnabled := FALSE;
FEnablePrevious := FALSE;
FResetRequested := TRUE;
FResetActive := TRUE;

IF Parent = 0 THEN
    EventPublisher.PublishEvent(Event := CreateFrameworkEvent(Name := AssertionName,
        ResourceName := ResourceName,
        State := E_State.Uninitialized,
        Severity := E_EventSeverity.Error,
        Message := 'Missing Test Case parent.'));
    RETURN;
END_IF;

ParentName := Parent.Name;
FullName := CONCAT(CONCAT(ParentName, '.'), AssertionName);
// SA0175: ASCII name contract; byte-based access is intentional and bounded.
{analysis -175}
FName := LEFT(FullName, UINT_TO_INT(GVL_Constants.NameLength));
{analysis +175}
FResourceName := ResourceName;
FObserveFirstCycle := ObserveFirstCycle;

IF NOT IsNameValid(Name := FullName, Depth := 4) THEN
    EventPublisher.PublishEvent(Event := CreateFrameworkEvent(Name := FName,
        ResourceName := FResourceName,
        State := E_State.Uninitialized,
        Severity := E_EventSeverity.Error,
        Message := CONCAT('Invalid Assertion name: ', FullName)));
    RETURN;
END_IF;

FInitialized := TRUE;
Initialize := TRUE;
END_METHOD

{region 'Documentation'}
(*!
<summary>TRUE after successful explicit initialization; retained by normal Reset.</summary>
*)
{endregion}
{attribute 'monitoring' := 'call'}
PROPERTY PUBLIC IsInitialized : BOOL //! TRUE after successful explicit initialization; retained by normal Reset.
GET // PUBLIC
IsInitialized := FInitialized;
END_GET
END_PROPERTY

{region 'Documentation'}
(*!
<summary>Length-limited hierarchical event name assigned by Initialize; retained by
Reset.</summary>
<description>

May contain an invalid diagnostic name; IsInitialized indicates validity.

</description>
*)
{endregion}
{attribute 'monitoring' := 'variable'}
PROPERTY PUBLIC Name : STRING(GVL_Constants.NameLength) //! Length-limited hierarchical event name assigned by Initialize; retained by Reset.
GET // PUBLIC
Name := FName;
END_GET
END_PROPERTY

{region 'Documentation'}
(*!
<summary>Indicate whether observation is enabled for the current accepted FB inputs.</summary>
<description>

Requires successful initialization, no reset in this call and Enabled. With
ObserveFirstCycle FALSE, a preceding enabled non-reset call is required. Overrides preserve
reset suppression and remain side-effect-free.

</description>
*)
{endregion}
{attribute 'monitoring' := 'call'}
PROPERTY PUBLIC ObservationActive : BOOL //! TRUE when initialized and enabled outside Reset, subject to the first-cycle setting and accepted call history.
GET // PUBLIC
ObservationActive := FInitialized AND NOT FResetActive AND FEnabled
    AND (FObserveFirstCycle OR FEnablePrevious);
END_GET
END_PROPERTY

{region 'Documentation'}
(*!
<summary>Read-only first-cycle setting supplied through Initialize; default TRUE, retained by
Reset.</summary>
<description>

Initialize with FALSE when the commanded test object must process before
observation.

</description>
*)
{endregion}
{attribute 'monitoring' := 'call'}
PROPERTY PUBLIC ObserveFirstCycle : BOOL //! Read-only first-cycle setting supplied through Initialize; default TRUE, retained by Reset.
GET // PUBLIC
ObserveFirstCycle := FObserveFirstCycle;
END_GET
END_PROPERTY

{region 'Documentation'}
(*!
<summary>Promote NotEvaluated to Passed without publishing a finding.</summary>
<description>

Leaves Passed, Failed and Error unchanged.

</description>
*)
{endregion}
METHOD PROTECTED Pass
IF FResult = E_Result.NotEvaluated THEN
    FResult := E_Result.Passed;
END_IF;
END_METHOD

{region 'Documentation'}
(*!
<summary>Request a reset to be consumed by the next FB call.</summary>
<description>

Does not immediately change Result. The consuming call clears result and observation
state and returns without checking; typed FB inputs must be bound for family-specific reset
work. Identity, settings and publisher are retained.

</description>
*)
{endregion}
METHOD PUBLIC Reset
FResetRequested := TRUE;
END_METHOD

{region 'Documentation'}
(*!
<summary>Reset family-specific observation state while FB inputs are bound.</summary>
<description>

The base implementation is empty. Override for owned history, snapshots or counters; do
not publish findings here. Called by the reset FB path, never directly by Initialize.

</description>
*)
{endregion}
METHOD PROTECTED ResetAssertion
END_METHOD

{region 'Documentation'}
(*!
<summary>Read-only tested resource context supplied through Initialize; default '', retained by
Reset.</summary>
*)
{endregion}
{attribute 'monitoring' := 'variable'}
PROPERTY PUBLIC ResourceName : STRING(GVL_Constants.ResourceNameLength) //! Read-only tested resource context supplied through Initialize; default '', retained by Reset.
GET // PUBLIC
ResourceName := FResourceName;
END_GET
END_PROPERTY

{region 'Documentation'}
(*!
<summary>Return the held assertion result.</summary>
<description>

Passed, Failed and Error do not de-escalate during checking. Consuming Reset or calling
Initialize clears the result to NotEvaluated. Disabled calls alone do not clear it.

</description>
*)
{endregion}
{attribute 'monitoring' := 'call'}
PROPERTY PUBLIC Result : E_Result //! Held assertion result; ordinary evaluation cannot lower Failed or Error.
GET // PUBLIC
Result := FResult;
END_GET
END_PROPERTY

END_FUNCTION_BLOCK

// ---- Framework/EventBuffer/POU/ResultEvents/CreateAssertionErrorEvent.TcPOU
{region 'Documentation'}
(*!
<summary>Constructs an assertion-error event without evaluating or publishing it.</summary>
<description>
The caller supplies the complete ASCII name, resource context and finding message.
</description>
*)
{endregion}
FUNCTION CreateAssertionErrorEvent : ST_Event //! Constructed event value; not published. The publisher assigns SequenceId and Timestamp.
VAR_INPUT
    Name : STRING(GVL_Constants.NameLength); //! Hierarchical owner name used to identify events; must satisfy the naming contract.
    ResourceName : STRING(GVL_Constants.ResourceNameLength) := ''; //! Optional resource context for diagnostics; empty by default.
    State : E_State; //! Owner lifecycle state recorded in the event.
    Message : STRING(GVL_Constants.MessageLength); //! Diagnostic text copied into the event within MessageLength.
END_VAR

CreateAssertionErrorEvent.SequenceId := 0;
CreateAssertionErrorEvent.Timestamp := 0;
CreateAssertionErrorEvent.OwnerScope := E_OwnerScope.Assertion;
CreateAssertionErrorEvent.EventType := E_EventType.Result;
CreateAssertionErrorEvent.Severity := SelectResultSeverity(Result := E_Result.Error);
CreateAssertionErrorEvent.Name := Name;
CreateAssertionErrorEvent.ResourceName := ResourceName;
CreateAssertionErrorEvent.State := State;
CreateAssertionErrorEvent.Result := E_Result.Error;
CreateAssertionErrorEvent.Message := Message;

END_FUNCTION

// ---- Framework/EventBuffer/POU/ResultEvents/CreateAssertionFailedEvent.TcPOU
{region 'Documentation'}
(*!
<summary>Constructs a failed-assertion event without evaluating or publishing it.</summary>
<description>
The caller supplies the complete ASCII name, resource context and finding message.
</description>
*)
{endregion}
FUNCTION CreateAssertionFailedEvent : ST_Event //! Constructed event value; not published. The publisher assigns SequenceId and Timestamp.
VAR_INPUT
    Name : STRING(GVL_Constants.NameLength); //! Hierarchical owner name used to identify events; must satisfy the naming contract.
    ResourceName : STRING(GVL_Constants.ResourceNameLength) := ''; //! Optional resource context for diagnostics; empty by default.
    State : E_State; //! Owner lifecycle state recorded in the event.
    Message : STRING(GVL_Constants.MessageLength); //! Diagnostic text copied into the event within MessageLength.
END_VAR

CreateAssertionFailedEvent.SequenceId := 0;
CreateAssertionFailedEvent.Timestamp := 0;
CreateAssertionFailedEvent.OwnerScope := E_OwnerScope.Assertion;
CreateAssertionFailedEvent.EventType := E_EventType.Result;
CreateAssertionFailedEvent.Severity := SelectResultSeverity(Result := E_Result.Failed);
CreateAssertionFailedEvent.Name := Name;
CreateAssertionFailedEvent.ResourceName := ResourceName;
CreateAssertionFailedEvent.State := State;
CreateAssertionFailedEvent.Result := E_Result.Failed;
CreateAssertionFailedEvent.Message := Message;

END_FUNCTION

// ---- SelfTests/TestSuites/TestSuite_Preparation.TcPOU
{region 'Documentation'}
(*!
<summary>Verifies Preparation status, resource actions and lifecycle handover in serial Test Cases.</summary>
*)
{endregion}
FUNCTION_BLOCK TestSuite_Preparation EXTENDS TestSuiteBase
VAR
    FInitialStatus : Test_PreparationInitialStatus;
    FStatusProjection : Test_PreparationStatusProjection;
    FDisabledObservation : Test_PreparationDisabledObservation;
    FReachesTarget : Test_PreparationReachesTarget;
    FDisableAndReenable : Test_PreparationDisableAndReenable;
    FCompletionTracksTarget : Test_PreparationCompletionTracksTarget;
    FResourceError : Test_PreparationResourceError;
    FMockInputs : Test_PreparationMockInputs;
    FTestCases : ARRAY[1..TestCaseCapacity] OF I_TestCase;
END_VAR
VAR CONSTANT
    TestCaseCapacity : UINT := 8;
END_VAR

SUPER^();

{region 'Documentation'}
(*!
<summary>Initializes all Preparation Test Cases and registers their deterministic serial order.</summary>
*)
{endregion}
METHOD PROTECTED Configure
VAR_IN_OUT
    // SA0167: Borrowed builder; VAR_IN_OUT creates no temporary instance.
    {attribute 'analysis' := '-167'}
    Builder : TestSuiteConfigurationBuilder; //! Borrowed owner configuration builder used only during this Configure call; register this owner's concrete children.
END_VAR
VAR
    TestConfig : ST_TestCaseConfig;
END_VAR
Builder.Initialize(Mode := E_OrchestrationMode.Serial,
    TestCases := FTestCases);

FInitialStatus.Initialize(Parent := THIS^,
    TestName := 'InitialStatus',
    Config := TestConfig);
Builder.Register(TestCase := FInitialStatus);

FStatusProjection.Initialize(Parent := THIS^,
    TestName := 'StatusProjection',
    Config := TestConfig);
Builder.Register(TestCase := FStatusProjection);

FDisabledObservation.Initialize(Parent := THIS^,
    TestName := 'DisabledObservation',
    Config := TestConfig);
Builder.Register(TestCase := FDisabledObservation);

FReachesTarget.Initialize(Parent := THIS^,
    TestName := 'ReachesTarget',
    Config := TestConfig);
Builder.Register(TestCase := FReachesTarget);

FDisableAndReenable.Initialize(Parent := THIS^,
    TestName := 'DisableAndReenable',
    Config := TestConfig);
Builder.Register(TestCase := FDisableAndReenable);

FCompletionTracksTarget.Initialize(Parent := THIS^,
    TestName := 'CompletionTracksTarget',
    Config := TestConfig);
Builder.Register(TestCase := FCompletionTracksTarget);

FResourceError.Initialize(Parent := THIS^,
    TestName := 'ResourceError',
    Config := TestConfig);
Builder.Register(TestCase := FResourceError);

FMockInputs.Initialize(Parent := THIS^,
    TestName := 'MockInputs',
    Config := TestConfig);
Builder.Register(TestCase := FMockInputs);
END_METHOD

{region 'Documentation'}
(*!
<summary>Returns the registered Test Case from the same array used during configuration.</summary>
*)
{endregion}
METHOD PUBLIC GetTestCase : I_TestCase //! Typed child interface at the original array index; zero when no entry is available.
VAR_INPUT
    Index : DINT; //! Original occupied child-array index, rather than an ordinal position.
END_VAR
GetTestCase := 0;
IF (ChildCount = 0) OR (Index < ChildArrayLowerBound)
    OR (DINT_TO_LINT(Index) >= DINT_TO_LINT(ChildArrayLowerBound) + UINT_TO_LINT(ChildCount)) THEN
    RETURN;
END_IF;

GetTestCase := FTestCases[Index];
END_METHOD

{region 'Documentation'}
(*!
<summary>Calls each owned Test Case once per initialized Suite cycle, including completion.</summary>
*)
{endregion}
METHOD PROTECTED ProcessTestCases
FInitialStatus();
FStatusProjection();
FDisabledObservation();
FReachesTarget();
FDisableAndReenable();
FCompletionTracksTarget();
FResourceError();
FMockInputs();
END_METHOD

END_FUNCTION_BLOCK

// ---- SelfTests/TestCases/TestSuite_Preparation/Test_PreparationInitialStatus.TcPOU
{region 'Documentation'}
(*!
<summary>Checks the untouched declaration snapshot through direct and interface reads; never calls the subject.</summary>
*)
{endregion}
FUNCTION_BLOCK Test_PreparationInitialStatus EXTENDS TestCaseBase
VAR
    FSubject : PreparationStatusProbe;
    FView : I_Preparation;
    FSnapshotCopy : ST_PreparationStatus;
    FObserved : ST_PreparationStatus;
    FExpected : ST_PreparationStatus;
    FObservedEnabled : BOOL;
    FExpectedEnabled : BOOL;
    FCheckPerformed : BOOL;
    FObservedCallCount : UDINT;
    FExpectedCallCount : UDINT;
    FCheckDiagnosticState : AssertEqual_Int;
    FCheckExecutionStatus : AssertEqual_Int;
    FCheckReady : AssertEqual_Bool;
    FCheckRunning : AssertEqual_Bool;
    FCheckCompleted : AssertEqual_Bool;
    FCheckError : AssertEqual_Bool;
    FCheckEnabled : AssertEqual_Bool;
    FCheckCallCount : AssertEqual_UDInt;
    FCheckCopyDetached : AssertEqual_Bool;
END_VAR
VAR CONSTANT
    DirectObservation : E_State := E_State.Running;
    DetachedSnapshot : E_State := E_State.Running + 1;
END_VAR

SUPER^();

{region 'Documentation'}
(*!
<summary>Contributes all owned Assertion results without executing the subjects.</summary>
*)
{endregion}
METHOD PROTECTED AggregateResults
VAR_INPUT
    Aggregator : I_ResultAggregator; //! Borrowed result sink owned by the outer Test Case; add this test's checking Assertions without resetting or retaining the sink.
END_VAR
Aggregator.AddProvider(Provider := FCheckDiagnosticState);
Aggregator.AddProvider(Provider := FCheckExecutionStatus);
Aggregator.AddProvider(Provider := FCheckReady);
Aggregator.AddProvider(Provider := FCheckRunning);
Aggregator.AddProvider(Provider := FCheckCompleted);
Aggregator.AddProvider(Provider := FCheckError);
Aggregator.AddProvider(Provider := FCheckEnabled);
Aggregator.AddProvider(Provider := FCheckCallCount);
Aggregator.AddProvider(Provider := FCheckCopyDetached);
END_METHOD

{region 'Documentation'}
(*!
<summary>Requires valid base configuration and every owned Assertion.</summary>
*)
{endregion}
METHOD PROTECTED CheckInitialization : BOOL //! TRUE when the inherited initialization check and this concrete fixture check both accept the setup.
CheckInitialization := FALSE;
IF NOT SUPER^.CheckInitialization() THEN
    RETURN;
END_IF;
IF NOT FCheckDiagnosticState.IsInitialized
    OR NOT FCheckExecutionStatus.IsInitialized
    OR NOT FCheckReady.IsInitialized
    OR NOT FCheckRunning.IsInitialized
    OR NOT FCheckCompleted.IsInitialized
    OR NOT FCheckError.IsInitialized
    OR NOT FCheckEnabled.IsInitialized
    OR NOT FCheckCallCount.IsInitialized
    OR NOT FCheckCopyDetached.IsInitialized THEN
    RETURN;
END_IF;

CheckInitialization := TRUE;
END_METHOD

{region 'Documentation'}
(*!
<summary>Configures this scenario, its local subjects and named Assertions.</summary>
*)
{endregion}
METHOD PROTECTED Configure
FPreparationStateCount := 0;
FTestStateCount := 2;
FCheckPerformed := FALSE;
FView := FSubject;
FSnapshotCopy.Completed := FALSE;

FCheckDiagnosticState.Initialize(Parent := THIS^,
    AssertionName := 'DiagnosticState');
FCheckExecutionStatus.Initialize(Parent := THIS^,
    AssertionName := 'ExecutionStatus');
FCheckReady.Initialize(Parent := THIS^,
    AssertionName := 'Ready');
FCheckRunning.Initialize(Parent := THIS^,
    AssertionName := 'Running');
FCheckCompleted.Initialize(Parent := THIS^,
    AssertionName := 'Completed');
FCheckError.Initialize(Parent := THIS^,
    AssertionName := 'Error');
FCheckEnabled.Initialize(Parent := THIS^,
    AssertionName := 'Enabled');
FCheckCallCount.Initialize(Parent := THIS^,
    AssertionName := 'CallCount');
FCheckCopyDetached.Initialize(Parent := THIS^,
    AssertionName := 'CopyDetached');
END_METHOD

{region 'Documentation'}
(*!
<summary>Ends scenario processing without issuing further resource commands.</summary>
*)
{endregion}
METHOD PROTECTED ProcessAbort
VAR_INPUT
    Enable : BOOL; //! Phase permission supplied by the owning Test Case; FALSE does not authorize progression, while observation may continue.
END_VAR
IF Enable THEN
    CompleteAbort();
END_IF;
END_METHOD

{region 'Documentation'}
(*!
<summary>Compares independent expected values with the captured observations; called when disabled as well.</summary>
*)
{endregion}
METHOD PROTECTED ProcessAssertions
VAR_INPUT
    Enable : BOOL; //! Phase permission supplied by the owning Test Case; FALSE does not authorize progression, while observation may continue.
END_VAR
FCheckDiagnosticState(Enable := Enable,
    State := State,
    IN := TO_INT(FObserved.State),
    Expected := TO_INT(FExpected.State));

FCheckExecutionStatus(Enable := Enable,
    State := State,
    IN := TO_INT(FObserved.ExecutionStatus),
    Expected := TO_INT(FExpected.ExecutionStatus));

FCheckReady(Enable := Enable,
    State := State,
    IN := FObserved.Ready,
    Expected := FExpected.Ready);

FCheckRunning(Enable := Enable,
    State := State,
    IN := FObserved.Running,
    Expected := FExpected.Running);

FCheckCompleted(Enable := Enable,
    State := State,
    IN := FObserved.Completed,
    Expected := FExpected.Completed);

FCheckError(Enable := Enable,
    State := State,
    IN := FObserved.Error,
    Expected := FExpected.Error);

FCheckEnabled(Enable := Enable,
    State := State,
    IN := FObservedEnabled,
    Expected := FExpectedEnabled);

FCheckCallCount(Enable := Enable,
    State := State,
    IN := FObservedCallCount,
    Expected := FExpectedCallCount);

FCheckCopyDetached(Enable := Enable,
    State := State,
    IN := FSnapshotCopy.Completed,
    Expected := State = DetachedSnapshot);

IF Enable
    AND FCheckDiagnosticState.EvaluationActive
    AND FCheckExecutionStatus.EvaluationActive
    AND FCheckReady.EvaluationActive
    AND FCheckRunning.EvaluationActive
    AND FCheckCompleted.EvaluationActive
    AND FCheckError.EvaluationActive
    AND FCheckEnabled.EvaluationActive
    AND FCheckCallCount.EvaluationActive
    AND FCheckCopyDetached.EvaluationActive THEN
    FCheckPerformed := TRUE;
END_IF;
END_METHOD

{region 'Documentation'}
(*!
<summary>Subjects are exercised by the test, not used as its start prerequisite.</summary>
*)
{endregion}
METHOD PROTECTED ProcessPreparations
VAR_INPUT
    // SA0033: Required hook; this scenario has no Preparation phase.
    {attribute 'analysis' := '-33'}
    Enable : BOOL; //! Phase permission supplied by the owning Test Case; FALSE does not authorize progression, while observation may continue.
END_VAR
END_METHOD

{region 'Documentation'}
(*!
<summary>Restores repeatable fixture state and resets Assertions before returning to Idle.</summary>
*)
{endregion}
METHOD PROTECTED ProcessReset
FCheckPerformed := FALSE;
FSnapshotCopy.Completed := FALSE;
FCheckDiagnosticState.Reset();
FCheckExecutionStatus.Reset();
FCheckReady.Reset();
FCheckRunning.Reset();
FCheckCompleted.Reset();
FCheckError.Reset();
FCheckEnabled.Reset();
FCheckCallCount.Reset();
FCheckCopyDetached.Reset();
CompleteReset();
END_METHOD

{region 'Documentation'}
(*!
<summary>Exercises one named scenario step per call; advances only after actual Assertion evaluation.</summary>
*)
{endregion}
METHOD PROTECTED ProcessTests
VAR_INPUT
    Enable : BOOL; //! Phase permission supplied by the owning Test Case; FALSE does not authorize progression, while observation may continue.
END_VAR
IF NOT Enable THEN
    RETURN;
END_IF;

IF FCheckPerformed THEN
    FCheckPerformed := FALSE;
    IF State = DetachedSnapshot THEN
        CompleteTests();
        RETURN;
    END_IF;
    NextTestState();
    IF NOT IsTestingActive THEN
        RETURN;
    END_IF;
END_IF;

CASE State OF
    DirectObservation:
        FObserved := FSubject.Status;
        FObservedEnabled := FSubject.Enabled;
        FExpected.State := E_State.Uninitialized;
        FExpected.ExecutionStatus := E_ExecutionStatus.Unknown;
        FExpected.Ready := FALSE;
        FExpected.Running := FALSE;
        FExpected.Completed := FALSE;
        FExpected.Error := FALSE;
        FExpectedEnabled := FALSE;
        FExpectedCallCount := 0;

    DetachedSnapshot:
        FSnapshotCopy := FView.Status;
        FSnapshotCopy.Completed := TRUE;
        FObserved := FView.Status;
        FObservedEnabled := FSubject.Enabled;
        FExpected.State := E_State.Uninitialized;
        FExpected.ExecutionStatus := E_ExecutionStatus.Unknown;
        FExpected.Ready := FALSE;
        FExpected.Running := FALSE;
        FExpected.Completed := FALSE;
        FExpected.Error := FALSE;
        FExpectedEnabled := FALSE;
        FExpectedCallCount := 0;

ELSE
    Error(Message := 'Unexpected Preparation test state.');
    RETURN;
END_CASE;

FObservedCallCount := FSubject.CallCount;
END_METHOD

END_FUNCTION_BLOCK

// ---- SelfTests/TestCases/TestSuite_Preparation/Helper/PreparationStatusProbe.TcPOU
{region 'Documentation'}
(*!
<summary>Exercises the real UpdateStatus mapping and counts Prepare calls without resource actions.</summary>
*)
{endregion}
FUNCTION_BLOCK PreparationStatusProbe EXTENDS PreparationBase
VAR_INPUT
    DiagnosticState : E_State := E_State.Idle; //! Scripted diagnostic state projected by Prepare.
    ExecutionStatus : E_ExecutionStatus := E_ExecutionStatus.Idle; //! Scripted execution classification projected by Prepare.
    Ready : BOOL := TRUE; //! Scripted readiness projected by Prepare.
END_VAR
VAR
    FCallCount : UDINT;
END_VAR

SUPER^();

{region 'Documentation'}
(*!
<summary>Current CallCount observation.</summary>
*)
{endregion}
{attribute 'monitoring' := 'call'}
PROPERTY PUBLIC CallCount : UDINT //! Current CallCount observation.
GET // PUBLIC
CallCount := FCallCount;
END_GET
END_PROPERTY

{region 'Documentation'}
(*!
<summary>Calls the inherited status projector once, including when disabled.</summary>
*)
{endregion}
METHOD PROTECTED Prepare
FCallCount := FCallCount + 1;
UpdateStatus(State := DiagnosticState,
    ExecutionStatus := ExecutionStatus,
    Ready := Ready);
END_METHOD

END_FUNCTION_BLOCK

// ---- Framework/Preparation/POU/PreparationBase.TcPOU
{region 'Documentation'}
(*!
<summary>Optional base for a resource Preparation controlled by level-based Enable.</summary>
<description>
Call SUPER^() once per task cycle. Implement Prepare to observe the resource on every call and
perform resource actions only while Enabled.

The base owns the accepted Enable view and status storage, not initialization, a reset
protocol, events or timeout supervision. The Test Case owns the Preparation timeout.

Disabled processing must not issue resource or cleanup commands. Removing Enable does not cancel
an already accepted resource command; the Test Case owns Reset/Abort handling.
</description>
*)
{endregion}
FUNCTION_BLOCK ABSTRACT PreparationBase IMPLEMENTS I_Preparation
VAR_INPUT
    Enable : BOOL; //! Permits resource-changing preparation work; disabled calls may still observe and report the resource.
END_VAR
VAR
    FEnabled : BOOL;
    /// Derived Prepare updates all applicable fields consistently with the Preparation contract.
    FStatus : ST_PreparationStatus;
END_VAR

FEnabled := Enable;
Prepare();

{region 'Documentation'}
(*!
<summary>Enable accepted at the last FB call; not proof of active resource manipulation.</summary>
*)
{endregion}
{attribute 'monitoring' := 'call'}
PROPERTY PUBLIC Enabled : BOOL //! Enable accepted at the last FB call; not proof of active resource manipulation.
GET // PUBLIC
Enabled := FEnabled;
END_GET
END_PROPERTY

{region 'Documentation'}
(*!
<summary>Observes the resource and maintains its Preparation status on every FB call.</summary>
<description>
This abstract hook has no base implementation to call. Use Enabled to gate resource-changing
work; disabled calls must still report current target, readiness and error observations.

On deactivation, stop resource manipulation and return any internal sequence to its executable
base state. Completed reports the current target condition, not a latched success. UpdateStatus may
be used to project consistent flags.
</description>
*)
{endregion}
METHOD PROTECTED ABSTRACT Prepare
END_METHOD

{region 'Documentation'}
(*!
<summary>Snapshot of the status maintained by the concrete Preparation.</summary>
*)
{endregion}
PROPERTY PUBLIC Status : ST_PreparationStatus //! Snapshot of the status maintained by the concrete Preparation.
GET // PUBLIC
Status := FStatus;
END_GET
END_PROPERTY

{region 'Documentation'}
(*!
<summary>Replaces the Preparation snapshot without performing resource work.</summary>
<description>
State is diagnostic context, independent of ExecutionStatus. Running, Completed and Error
follow ExecutionStatus; Ready is suppressed only while Running.

Select E_ExecutionStatus.Idle only when Ready is TRUE and neither work, completion nor error applies; otherwise
select E_ExecutionStatus.NotReady. This method does not validate that choice, latch completion, publish events or
supervise timeouts.
</description>
*)
{endregion}
METHOD PROTECTED UpdateStatus
VAR_INPUT
    State : E_State; //! Concrete Preparation's lifecycle state; independent of the execution-status classification.
    ExecutionStatus : E_ExecutionStatus; //! Execution classification used to derive Running, Completed and Error in the Preparation snapshot.
    Ready : BOOL; //! Resource can be driven to the target state; suppressed while Running. Does not mean target reached.
END_VAR
FStatus.State := State;
FStatus.ExecutionStatus := ExecutionStatus;
FStatus.Running := ExecutionStatus = E_ExecutionStatus.Running;
FStatus.Completed := ExecutionStatus = E_ExecutionStatus.Completed;
FStatus.Error := ExecutionStatus = E_ExecutionStatus.Error;
FStatus.Ready := Ready AND NOT FStatus.Running;
END_METHOD

END_FUNCTION_BLOCK

// ---- Framework/Assertions/POU/BasicTypes/Int/AssertEqual_Int.TcPOU
{region 'Documentation'}
(*!
<summary>Checks equality with the expected INT value.</summary>
*)
{endregion}
FUNCTION_BLOCK AssertEqual_Int EXTENDS AssertionBase
VAR_INPUT
    IN : INT; //! Actual value checked or observed by this Assertion.
    Expected : INT; //! Reference value for comparison with IN.
END_VAR

SUPER^();

{region 'Documentation'}
(*!
<summary>Check equality with the expected INT value.</summary>
*)
{endregion}
METHOD PROTECTED Assert
VAR
    Message : STRING(GVL_Constants.MessageLength);
    ExpectedText : STRING(GVL_Constants.AssertionValueLength);
    ActualText : STRING(GVL_Constants.AssertionValueLength);
END_VAR
IF NOT EvaluationActive THEN
    RETURN;
END_IF;

IF Result = E_Result.Error THEN
    RETURN;
END_IF;

IF Result = E_Result.Failed THEN
    RETURN;
END_IF;

IF IN <> Expected THEN
    ExpectedText := INT_TO_STRING(Expected);
    ActualText := INT_TO_STRING(IN);
    Message := CONCAT('Assertion failed: values are not equal. Expected = ',
        ExpectedText);
    Message := CONCAT(Message, ', Actual = ');
    Message := CONCAT(Message, ActualText);
    Message := CONCAT(Message, '.');
    Fail(Message := Message);
    RETURN;
END_IF;

Pass();
END_METHOD

END_FUNCTION_BLOCK

// ---- Framework/Assertions/POU/BasicTypes/Bool/AssertEqual_Bool.TcPOU
{region 'Documentation'}
(*!
<summary>Checks equality with the expected BOOL value.</summary>
*)
{endregion}
FUNCTION_BLOCK AssertEqual_Bool EXTENDS AssertionBase
VAR_INPUT
    IN : BOOL; //! Actual value checked or observed by this Assertion.
    Expected : BOOL; //! Reference value for comparison with IN.
END_VAR

SUPER^();

{region 'Documentation'}
(*!
<summary>Check equality with the expected BOOL value.</summary>
*)
{endregion}
METHOD PROTECTED Assert
VAR
    Message : STRING(GVL_Constants.MessageLength);
    ExpectedText : STRING(GVL_Constants.AssertionValueLength);
    ActualText : STRING(GVL_Constants.AssertionValueLength);
END_VAR
IF NOT EvaluationActive THEN
    RETURN;
END_IF;

IF Result = E_Result.Error THEN
    RETURN;
END_IF;

IF Result = E_Result.Failed THEN
    RETURN;
END_IF;

IF IN <> Expected THEN
    ExpectedText := BOOL_TO_STRING(Expected);
    ActualText := BOOL_TO_STRING(IN);
    Message := CONCAT('Assertion failed: values are not equal. Expected = ',
        ExpectedText);
    Message := CONCAT(Message, ', Actual = ');
    Message := CONCAT(Message, ActualText);
    Message := CONCAT(Message, '.');
    Fail(Message := Message);
    RETURN;
END_IF;

Pass();
END_METHOD

END_FUNCTION_BLOCK

// ---- SelfTests/TestCases/TestSuite_Preparation/Test_PreparationStatusProjection.TcPOU
{region 'Documentation'}
(*!
<summary>Checks real status projection, independent diagnostic state, flag replacement and Prepare invocation count.</summary>
*)
{endregion}
FUNCTION_BLOCK Test_PreparationStatusProjection EXTENDS TestCaseBase
VAR
    FSubject : PreparationStatusProbe;
    FView : I_Preparation;
    FInitialCallCount : UDINT;
    FObserved : ST_PreparationStatus;
    FExpected : ST_PreparationStatus;
    FObservedEnabled : BOOL;
    FExpectedEnabled : BOOL;
    FCheckPerformed : BOOL;
    FObservedCallCount : UDINT;
    FExpectedCallCount : UDINT;
    FCheckDiagnosticState : AssertEqual_Int;
    FCheckExecutionStatus : AssertEqual_Int;
    FCheckReady : AssertEqual_Bool;
    FCheckRunning : AssertEqual_Bool;
    FCheckCompleted : AssertEqual_Bool;
    FCheckError : AssertEqual_Bool;
    FCheckEnabled : AssertEqual_Bool;
    FCheckCallCount : AssertEqual_UDInt;
END_VAR
VAR CONSTANT
    IdleObservation : E_State := E_State.Running;
    UnavailableObservation : E_State := E_State.Running + 1;
    RunningObservation : E_State := E_State.Running + 2;
    IndependentDiagnosticState : E_State := E_State.Running + 3;
    ErrorObservation : E_State := E_State.Running + 4;
    ClearedFlags : E_State := E_State.Running + 5;
END_VAR

SUPER^();

{region 'Documentation'}
(*!
<summary>Contributes all owned Assertion results without executing the subjects.</summary>
*)
{endregion}
METHOD PROTECTED AggregateResults
VAR_INPUT
    Aggregator : I_ResultAggregator; //! Borrowed result sink owned by the outer Test Case; add this test's checking Assertions without resetting or retaining the sink.
END_VAR
Aggregator.AddProvider(Provider := FCheckDiagnosticState);
Aggregator.AddProvider(Provider := FCheckExecutionStatus);
Aggregator.AddProvider(Provider := FCheckReady);
Aggregator.AddProvider(Provider := FCheckRunning);
Aggregator.AddProvider(Provider := FCheckCompleted);
Aggregator.AddProvider(Provider := FCheckError);
Aggregator.AddProvider(Provider := FCheckEnabled);
Aggregator.AddProvider(Provider := FCheckCallCount);
END_METHOD

{region 'Documentation'}
(*!
<summary>Requires valid base configuration and every owned Assertion.</summary>
*)
{endregion}
METHOD PROTECTED CheckInitialization : BOOL //! TRUE when the inherited initialization check and this concrete fixture check both accept the setup.
CheckInitialization := FALSE;
IF NOT SUPER^.CheckInitialization() THEN
    RETURN;
END_IF;
IF NOT FCheckDiagnosticState.IsInitialized
    OR NOT FCheckExecutionStatus.IsInitialized
    OR NOT FCheckReady.IsInitialized
    OR NOT FCheckRunning.IsInitialized
    OR NOT FCheckCompleted.IsInitialized
    OR NOT FCheckError.IsInitialized
    OR NOT FCheckEnabled.IsInitialized
    OR NOT FCheckCallCount.IsInitialized THEN
    RETURN;
END_IF;

CheckInitialization := TRUE;
END_METHOD

{region 'Documentation'}
(*!
<summary>Configures this scenario, its local subjects and named Assertions.</summary>
*)
{endregion}
METHOD PROTECTED Configure
FPreparationStateCount := 0;
FTestStateCount := 6;
FCheckPerformed := FALSE;
FView := FSubject;
FInitialCallCount := FSubject.CallCount;

FCheckDiagnosticState.Initialize(Parent := THIS^,
    AssertionName := 'DiagnosticState');
FCheckExecutionStatus.Initialize(Parent := THIS^,
    AssertionName := 'ExecutionStatus');
FCheckReady.Initialize(Parent := THIS^,
    AssertionName := 'Ready');
FCheckRunning.Initialize(Parent := THIS^,
    AssertionName := 'Running');
FCheckCompleted.Initialize(Parent := THIS^,
    AssertionName := 'Completed');
FCheckError.Initialize(Parent := THIS^,
    AssertionName := 'Error');
FCheckEnabled.Initialize(Parent := THIS^,
    AssertionName := 'Enabled');
FCheckCallCount.Initialize(Parent := THIS^,
    AssertionName := 'CallCount');
END_METHOD

{region 'Documentation'}
(*!
<summary>Ends scenario processing without issuing further resource commands.</summary>
*)
{endregion}
METHOD PROTECTED ProcessAbort
VAR_INPUT
    Enable : BOOL; //! Phase permission supplied by the owning Test Case; FALSE does not authorize progression, while observation may continue.
END_VAR
IF Enable THEN
    CompleteAbort();
END_IF;
END_METHOD

{region 'Documentation'}
(*!
<summary>Compares independent expected values with the captured observations; called when disabled as well.</summary>
*)
{endregion}
METHOD PROTECTED ProcessAssertions
VAR_INPUT
    Enable : BOOL; //! Phase permission supplied by the owning Test Case; FALSE does not authorize progression, while observation may continue.
END_VAR
FCheckDiagnosticState(Enable := Enable,
    State := State,
    IN := TO_INT(FObserved.State),
    Expected := TO_INT(FExpected.State));

FCheckExecutionStatus(Enable := Enable,
    State := State,
    IN := TO_INT(FObserved.ExecutionStatus),
    Expected := TO_INT(FExpected.ExecutionStatus));

FCheckReady(Enable := Enable,
    State := State,
    IN := FObserved.Ready,
    Expected := FExpected.Ready);

FCheckRunning(Enable := Enable,
    State := State,
    IN := FObserved.Running,
    Expected := FExpected.Running);

FCheckCompleted(Enable := Enable,
    State := State,
    IN := FObserved.Completed,
    Expected := FExpected.Completed);

FCheckError(Enable := Enable,
    State := State,
    IN := FObserved.Error,
    Expected := FExpected.Error);

FCheckEnabled(Enable := Enable,
    State := State,
    IN := FObservedEnabled,
    Expected := FExpectedEnabled);

FCheckCallCount(Enable := Enable,
    State := State,
    IN := FObservedCallCount,
    Expected := FExpectedCallCount);

IF Enable
    AND FCheckDiagnosticState.EvaluationActive
    AND FCheckExecutionStatus.EvaluationActive
    AND FCheckReady.EvaluationActive
    AND FCheckRunning.EvaluationActive
    AND FCheckCompleted.EvaluationActive
    AND FCheckError.EvaluationActive
    AND FCheckEnabled.EvaluationActive
    AND FCheckCallCount.EvaluationActive THEN
    FCheckPerformed := TRUE;
END_IF;
END_METHOD

{region 'Documentation'}
(*!
<summary>Subjects are exercised by the test, not used as its start prerequisite.</summary>
*)
{endregion}
METHOD PROTECTED ProcessPreparations
VAR_INPUT
    // SA0033: Required hook; this scenario has no Preparation phase.
    {attribute 'analysis' := '-33'}
    Enable : BOOL; //! Phase permission supplied by the owning Test Case; FALSE does not authorize progression, while observation may continue.
END_VAR
END_METHOD

{region 'Documentation'}
(*!
<summary>Restores repeatable fixture state and resets Assertions before returning to Idle.</summary>
*)
{endregion}
METHOD PROTECTED ProcessReset
FCheckPerformed := FALSE;
FInitialCallCount := FSubject.CallCount;
FCheckDiagnosticState.Reset();
FCheckExecutionStatus.Reset();
FCheckReady.Reset();
FCheckRunning.Reset();
FCheckCompleted.Reset();
FCheckError.Reset();
FCheckEnabled.Reset();
FCheckCallCount.Reset();
CompleteReset();
END_METHOD

{region 'Documentation'}
(*!
<summary>Exercises one named scenario step per call; advances only after actual Assertion evaluation.</summary>
*)
{endregion}
METHOD PROTECTED ProcessTests
VAR_INPUT
    Enable : BOOL; //! Phase permission supplied by the owning Test Case; FALSE does not authorize progression, while observation may continue.
END_VAR
IF NOT Enable THEN
    RETURN;
END_IF;

IF FCheckPerformed THEN
    FCheckPerformed := FALSE;
    IF State = ClearedFlags THEN
        CompleteTests();
        RETURN;
    END_IF;
    NextTestState();
    IF NOT IsTestingActive THEN
        RETURN;
    END_IF;
END_IF;

CASE State OF
    IdleObservation:
        FSubject(Enable := FALSE,
            DiagnosticState := E_State.Idle,
            ExecutionStatus := E_ExecutionStatus.Idle,
            Ready := TRUE);
        FExpected.State := E_State.Idle;
        FExpected.ExecutionStatus := E_ExecutionStatus.Idle;
        FExpected.Ready := TRUE;
        FExpected.Running := FALSE;
        FExpected.Completed := FALSE;
        FExpected.Error := FALSE;
        FExpectedEnabled := FALSE;
        FExpectedCallCount := 1;

    UnavailableObservation:
        FSubject(Enable := TRUE,
            DiagnosticState := E_State.Idle,
            ExecutionStatus := E_ExecutionStatus.NotReady,
            Ready := FALSE);
        FExpected.State := E_State.Idle;
        FExpected.ExecutionStatus := E_ExecutionStatus.NotReady;
        FExpected.Ready := FALSE;
        FExpected.Running := FALSE;
        FExpected.Completed := FALSE;
        FExpected.Error := FALSE;
        FExpectedEnabled := TRUE;
        FExpectedCallCount := 2;

    RunningObservation:
        FSubject(Enable := TRUE,
            DiagnosticState := E_State.Preparing,
            ExecutionStatus := E_ExecutionStatus.Running,
            Ready := TRUE);
        FExpected.State := E_State.Preparing;
        FExpected.ExecutionStatus := E_ExecutionStatus.Running;
        FExpected.Ready := FALSE;
        FExpected.Running := TRUE;
        FExpected.Completed := FALSE;
        FExpected.Error := FALSE;
        FExpectedEnabled := TRUE;
        FExpectedCallCount := 3;

    IndependentDiagnosticState:
        FSubject(Enable := FALSE,
            DiagnosticState := E_State.Idle,
            ExecutionStatus := E_ExecutionStatus.Completed,
            Ready := TRUE);
        FExpected.State := E_State.Idle;
        FExpected.ExecutionStatus := E_ExecutionStatus.Completed;
        FExpected.Ready := TRUE;
        FExpected.Running := FALSE;
        FExpected.Completed := TRUE;
        FExpected.Error := FALSE;
        FExpectedEnabled := FALSE;
        FExpectedCallCount := 4;

    ErrorObservation:
        FSubject(Enable := FALSE,
            DiagnosticState := E_State.Error,
            ExecutionStatus := E_ExecutionStatus.Error,
            Ready := TRUE);
        FExpected.State := E_State.Error;
        FExpected.ExecutionStatus := E_ExecutionStatus.Error;
        FExpected.Ready := TRUE;
        FExpected.Running := FALSE;
        FExpected.Completed := FALSE;
        FExpected.Error := TRUE;
        FExpectedEnabled := FALSE;
        FExpectedCallCount := 5;

    ClearedFlags:
        FSubject(Enable := TRUE,
            DiagnosticState := E_State.Idle,
            ExecutionStatus := E_ExecutionStatus.Idle,
            Ready := TRUE);
        FExpected.State := E_State.Idle;
        FExpected.ExecutionStatus := E_ExecutionStatus.Idle;
        FExpected.Ready := TRUE;
        FExpected.Running := FALSE;
        FExpected.Completed := FALSE;
        FExpected.Error := FALSE;
        FExpectedEnabled := TRUE;
        FExpectedCallCount := 6;

ELSE
    Error(Message := 'Unexpected Preparation test state.');
    RETURN;
END_CASE;

FObserved := FView.Status;
FObservedEnabled := FSubject.Enabled;

FObservedCallCount := FSubject.CallCount - FInitialCallCount;
END_METHOD

END_FUNCTION_BLOCK

// ---- SelfTests/TestCases/TestSuite_Preparation/Test_PreparationDisabledObservation.TcPOU
{region 'Documentation'}
(*!
<summary>Checks disabled observation, absence of command writes and current completion after externally driven resource changes.</summary>
*)
{endregion}
FUNCTION_BLOCK Test_PreparationDisabledObservation EXTENDS TestCaseBase
VAR
    FSubject : Prepare_ValueAtTarget;
    FResource : PreparationResource;
    FView : I_Preparation;
    FObserved : ST_PreparationStatus;
    FExpected : ST_PreparationStatus;
    FObservedEnabled : BOOL;
    FExpectedEnabled : BOOL;
    FCheckPerformed : BOOL;
    FObservedCommandWrites : UDINT;
    FExpectedCommandWrites : UDINT;
    FObservedActualValue : DINT;
    FExpectedActualValue : DINT;
    FObservedRequestedValue : DINT;
    FExpectedRequestedValue : DINT;
    FCheckDiagnosticState : AssertEqual_Int;
    FCheckExecutionStatus : AssertEqual_Int;
    FCheckReady : AssertEqual_Bool;
    FCheckRunning : AssertEqual_Bool;
    FCheckCompleted : AssertEqual_Bool;
    FCheckError : AssertEqual_Bool;
    FCheckEnabled : AssertEqual_Bool;
    FCheckCommandWrites : AssertEqual_UDInt;
    FCheckActualValue : AssertEqual_DInt;
    FCheckRequestedValue : AssertEqual_DInt;
END_VAR
VAR CONSTANT
    ReadyObservation : E_State := E_State.Running;
    NotReadyObservation : E_State := E_State.Running + 1;
    ExternalMovement : E_State := E_State.Running + 2;
    TargetObservation : E_State := E_State.Running + 3;
    TargetDeparture : E_State := E_State.Running + 4;
    UnsupportedCondition : E_State := E_State.Running + 5;
    FaultObservation : E_State := E_State.Running + 6;
    RecoveryObservation : E_State := E_State.Running + 7;
END_VAR

SUPER^();

{region 'Documentation'}
(*!
<summary>Contributes all owned Assertion results without executing the subjects.</summary>
*)
{endregion}
METHOD PROTECTED AggregateResults
VAR_INPUT
    Aggregator : I_ResultAggregator; //! Borrowed result sink owned by the outer Test Case; add this test's checking Assertions without resetting or retaining the sink.
END_VAR
Aggregator.AddProvider(Provider := FCheckDiagnosticState);
Aggregator.AddProvider(Provider := FCheckExecutionStatus);
Aggregator.AddProvider(Provider := FCheckReady);
Aggregator.AddProvider(Provider := FCheckRunning);
Aggregator.AddProvider(Provider := FCheckCompleted);
Aggregator.AddProvider(Provider := FCheckError);
Aggregator.AddProvider(Provider := FCheckEnabled);
Aggregator.AddProvider(Provider := FCheckCommandWrites);
Aggregator.AddProvider(Provider := FCheckActualValue);
Aggregator.AddProvider(Provider := FCheckRequestedValue);
END_METHOD

{region 'Documentation'}
(*!
<summary>Requires valid base configuration and every owned Assertion.</summary>
*)
{endregion}
METHOD PROTECTED CheckInitialization : BOOL //! TRUE when the inherited initialization check and this concrete fixture check both accept the setup.
CheckInitialization := FALSE;
IF NOT SUPER^.CheckInitialization() THEN
    RETURN;
END_IF;
IF NOT FCheckDiagnosticState.IsInitialized
    OR NOT FCheckExecutionStatus.IsInitialized
    OR NOT FCheckReady.IsInitialized
    OR NOT FCheckRunning.IsInitialized
    OR NOT FCheckCompleted.IsInitialized
    OR NOT FCheckError.IsInitialized
    OR NOT FCheckEnabled.IsInitialized
    OR NOT FCheckCommandWrites.IsInitialized
    OR NOT FCheckActualValue.IsInitialized
    OR NOT FCheckRequestedValue.IsInitialized THEN
    RETURN;
END_IF;

CheckInitialization := TRUE;
END_METHOD

{region 'Documentation'}
(*!
<summary>Configures this scenario, its local subjects and named Assertions.</summary>
*)
{endregion}
METHOD PROTECTED Configure
FPreparationStateCount := 0;
FTestStateCount := 8;
FCheckPerformed := FALSE;
FResource.Initialize(InitialValue := 2);
FSubject.Initialize(Resource := FResource);
FView := FSubject;

FCheckDiagnosticState.Initialize(Parent := THIS^,
    AssertionName := 'DiagnosticState');
FCheckExecutionStatus.Initialize(Parent := THIS^,
    AssertionName := 'ExecutionStatus');
FCheckReady.Initialize(Parent := THIS^,
    AssertionName := 'Ready');
FCheckRunning.Initialize(Parent := THIS^,
    AssertionName := 'Running');
FCheckCompleted.Initialize(Parent := THIS^,
    AssertionName := 'Completed');
FCheckError.Initialize(Parent := THIS^,
    AssertionName := 'Error');
FCheckEnabled.Initialize(Parent := THIS^,
    AssertionName := 'Enabled');
FCheckCommandWrites.Initialize(Parent := THIS^,
    AssertionName := 'CommandWrites');
FCheckActualValue.Initialize(Parent := THIS^,
    AssertionName := 'ActualValue');
FCheckRequestedValue.Initialize(Parent := THIS^,
    AssertionName := 'RequestedValue');
END_METHOD

{region 'Documentation'}
(*!
<summary>Ends scenario processing without issuing further resource commands.</summary>
*)
{endregion}
METHOD PROTECTED ProcessAbort
VAR_INPUT
    Enable : BOOL; //! Phase permission supplied by the owning Test Case; FALSE does not authorize progression, while observation may continue.
END_VAR
IF Enable THEN
    CompleteAbort();
END_IF;
END_METHOD

{region 'Documentation'}
(*!
<summary>Compares independent expected values with the captured observations; called when disabled as well.</summary>
*)
{endregion}
METHOD PROTECTED ProcessAssertions
VAR_INPUT
    Enable : BOOL; //! Phase permission supplied by the owning Test Case; FALSE does not authorize progression, while observation may continue.
END_VAR
FCheckDiagnosticState(Enable := Enable,
    State := State,
    IN := TO_INT(FObserved.State),
    Expected := TO_INT(FExpected.State));

FCheckExecutionStatus(Enable := Enable,
    State := State,
    IN := TO_INT(FObserved.ExecutionStatus),
    Expected := TO_INT(FExpected.ExecutionStatus));

FCheckReady(Enable := Enable,
    State := State,
    IN := FObserved.Ready,
    Expected := FExpected.Ready);

FCheckRunning(Enable := Enable,
    State := State,
    IN := FObserved.Running,
    Expected := FExpected.Running);

FCheckCompleted(Enable := Enable,
    State := State,
    IN := FObserved.Completed,
    Expected := FExpected.Completed);

FCheckError(Enable := Enable,
    State := State,
    IN := FObserved.Error,
    Expected := FExpected.Error);

FCheckEnabled(Enable := Enable,
    State := State,
    IN := FObservedEnabled,
    Expected := FExpectedEnabled);

FCheckCommandWrites(Enable := Enable,
    State := State,
    IN := FObservedCommandWrites,
    Expected := FExpectedCommandWrites);

FCheckActualValue(Enable := Enable,
    State := State,
    IN := FObservedActualValue,
    Expected := FExpectedActualValue);

FCheckRequestedValue(Enable := Enable,
    State := State,
    IN := FObservedRequestedValue,
    Expected := FExpectedRequestedValue);

IF Enable
    AND FCheckDiagnosticState.EvaluationActive
    AND FCheckExecutionStatus.EvaluationActive
    AND FCheckReady.EvaluationActive
    AND FCheckRunning.EvaluationActive
    AND FCheckCompleted.EvaluationActive
    AND FCheckError.EvaluationActive
    AND FCheckEnabled.EvaluationActive
    AND FCheckCommandWrites.EvaluationActive
    AND FCheckActualValue.EvaluationActive
    AND FCheckRequestedValue.EvaluationActive THEN
    FCheckPerformed := TRUE;
END_IF;
END_METHOD

{region 'Documentation'}
(*!
<summary>Subjects are exercised by the test, not used as its start prerequisite.</summary>
*)
{endregion}
METHOD PROTECTED ProcessPreparations
VAR_INPUT
    // SA0033: Required hook; this scenario has no Preparation phase.
    {attribute 'analysis' := '-33'}
    Enable : BOOL; //! Phase permission supplied by the owning Test Case; FALSE does not authorize progression, while observation may continue.
END_VAR
END_METHOD

{region 'Documentation'}
(*!
<summary>Restores repeatable fixture state and resets Assertions before returning to Idle.</summary>
*)
{endregion}
METHOD PROTECTED ProcessReset
FCheckPerformed := FALSE;
FResource.Initialize(InitialValue := 2);
FSubject.Initialize(Resource := FResource);
FView := FSubject;
FCheckDiagnosticState.Reset();
FCheckExecutionStatus.Reset();
FCheckReady.Reset();
FCheckRunning.Reset();
FCheckCompleted.Reset();
FCheckError.Reset();
FCheckEnabled.Reset();
FCheckCommandWrites.Reset();
FCheckActualValue.Reset();
FCheckRequestedValue.Reset();
CompleteReset();
END_METHOD

{region 'Documentation'}
(*!
<summary>Exercises one named scenario step per call; advances only after actual Assertion evaluation.</summary>
*)
{endregion}
METHOD PROTECTED ProcessTests
VAR_INPUT
    Enable : BOOL; //! Phase permission supplied by the owning Test Case; FALSE does not authorize progression, while observation may continue.
END_VAR
IF NOT Enable THEN
    RETURN;
END_IF;

IF FCheckPerformed THEN
    FCheckPerformed := FALSE;
    IF State = RecoveryObservation THEN
        CompleteTests();
        RETURN;
    END_IF;
    NextTestState();
    IF NOT IsTestingActive THEN
        RETURN;
    END_IF;
END_IF;

CASE State OF
    ReadyObservation:
        FResource(Available := TRUE,
            Fault := FALSE,
            Advance := TRUE);
        FSubject(Enable := FALSE,
            TargetValue := 0);
        FExpected.State := E_State.Idle;
        FExpected.ExecutionStatus := E_ExecutionStatus.Idle;
        FExpected.Ready := TRUE;
        FExpected.Running := FALSE;
        FExpected.Completed := FALSE;
        FExpected.Error := FALSE;
        FExpectedEnabled := FALSE;
        FExpectedCommandWrites := 0;
        FExpectedActualValue := 2;
        FExpectedRequestedValue := 2;

    NotReadyObservation:
        FResource(Available := FALSE,
            Fault := FALSE,
            Advance := TRUE);
        FSubject(Enable := FALSE,
            TargetValue := 0);
        FExpected.State := E_State.Idle;
        FExpected.ExecutionStatus := E_ExecutionStatus.NotReady;
        FExpected.Ready := FALSE;
        FExpected.Running := FALSE;
        FExpected.Completed := FALSE;
        FExpected.Error := FALSE;
        FExpectedEnabled := FALSE;
        FExpectedCommandWrites := 0;
        FExpectedActualValue := 2;
        FExpectedRequestedValue := 2;

    ExternalMovement:
        FResource.RequestValue(Value := 0);
        FResource(Available := TRUE,
            Fault := FALSE,
            Advance := TRUE);
        FSubject(Enable := FALSE,
            TargetValue := 0);
        FExpected.State := E_State.Idle;
        FExpected.ExecutionStatus := E_ExecutionStatus.Idle;
        FExpected.Ready := TRUE;
        FExpected.Running := FALSE;
        FExpected.Completed := FALSE;
        FExpected.Error := FALSE;
        FExpectedEnabled := FALSE;
        FExpectedCommandWrites := 1;
        FExpectedActualValue := 1;
        FExpectedRequestedValue := 0;

    TargetObservation:
        FResource(Available := TRUE,
            Fault := FALSE,
            Advance := TRUE);
        FSubject(Enable := FALSE,
            TargetValue := 0);
        FExpected.State := E_State.Completed;
        FExpected.ExecutionStatus := E_ExecutionStatus.Completed;
        FExpected.Ready := TRUE;
        FExpected.Running := FALSE;
        FExpected.Completed := TRUE;
        FExpected.Error := FALSE;
        FExpectedEnabled := FALSE;
        FExpectedCommandWrites := 1;
        FExpectedActualValue := 0;
        FExpectedRequestedValue := 0;

    TargetDeparture:
        FResource.RequestValue(Value := 2);
        FResource(Available := TRUE,
            Fault := FALSE,
            Advance := TRUE);
        FSubject(Enable := FALSE,
            TargetValue := 0);
        FExpected.State := E_State.Idle;
        FExpected.ExecutionStatus := E_ExecutionStatus.Idle;
        FExpected.Ready := TRUE;
        FExpected.Running := FALSE;
        FExpected.Completed := FALSE;
        FExpected.Error := FALSE;
        FExpectedEnabled := FALSE;
        FExpectedCommandWrites := 2;
        FExpectedActualValue := 1;
        FExpectedRequestedValue := 2;

    UnsupportedCondition:
        FResource(Available := FALSE,
            Fault := FALSE,
            Advance := TRUE);
        FSubject(Enable := FALSE,
            TargetValue := 0);
        FExpected.State := E_State.Idle;
        FExpected.ExecutionStatus := E_ExecutionStatus.NotReady;
        FExpected.Ready := FALSE;
        FExpected.Running := FALSE;
        FExpected.Completed := FALSE;
        FExpected.Error := FALSE;
        FExpectedEnabled := FALSE;
        FExpectedCommandWrites := 2;
        FExpectedActualValue := 1;
        FExpectedRequestedValue := 2;

    FaultObservation:
        FResource(Available := TRUE,
            Fault := TRUE,
            Advance := TRUE);
        FSubject(Enable := FALSE,
            TargetValue := 0);
        FExpected.State := E_State.Error;
        FExpected.ExecutionStatus := E_ExecutionStatus.Error;
        FExpected.Ready := FALSE;
        FExpected.Running := FALSE;
        FExpected.Completed := FALSE;
        FExpected.Error := TRUE;
        FExpectedEnabled := FALSE;
        FExpectedCommandWrites := 2;
        FExpectedActualValue := 1;
        FExpectedRequestedValue := 2;

    RecoveryObservation:
        FResource(Available := TRUE,
            Fault := FALSE,
            Advance := FALSE);
        FSubject(Enable := FALSE,
            TargetValue := 0);
        FExpected.State := E_State.Idle;
        FExpected.ExecutionStatus := E_ExecutionStatus.Idle;
        FExpected.Ready := TRUE;
        FExpected.Running := FALSE;
        FExpected.Completed := FALSE;
        FExpected.Error := FALSE;
        FExpectedEnabled := FALSE;
        FExpectedCommandWrites := 2;
        FExpectedActualValue := 1;
        FExpectedRequestedValue := 2;

ELSE
    Error(Message := 'Unexpected Preparation test state.');
    RETURN;
END_CASE;

FObserved := FView.Status;
FObservedEnabled := FSubject.Enabled;

FObservedCommandWrites := FResource.CommandWriteCount;
FObservedActualValue := FResource.ActualValue;
FObservedRequestedValue := FResource.RequestedValue;
END_METHOD

END_FUNCTION_BLOCK

// ---- SelfTests/TestCases/TestSuite_Preparation/Helper/Prepare_ValueAtTarget.TcPOU
{region 'Documentation'}
(*!
<summary>Establishes both request and feedback at TargetValue using the real PreparationBase status projection. The test owns and calls the resource separately. Disabled calls observe without commands or cancellation.</summary>
*)
{endregion}
FUNCTION_BLOCK Prepare_ValueAtTarget EXTENDS PreparationBase
VAR_INPUT
    TargetValue : DINT := 0; //! Requested resource value while enabled; disabled calls observe without issuing commands.
END_VAR
VAR
    FResource : REFERENCE TO PreparationResource;
END_VAR

SUPER^();

{region 'Documentation'}
(*!
<summary>Binds the test-owned resource before use. Its lifetime must cover all Preparation calls. No resource access or feedback change; subsequent FB calls refresh the inherited observation.</summary>
*)
{endregion}
METHOD PUBLIC Initialize
VAR_IN_OUT
    // SA0167: Borrowed static resource, not a temporary FB instance.
    {attribute 'analysis' := '-167'}
    Resource : PreparationResource; //! Borrowed static resource retained by reference; keep it alive and stable for all preparation calls.
END_VAR
FResource REF= Resource;
END_METHOD

{region 'Documentation'}
(*!
<summary>Observes every call; errors and unsupported resource conditions prevent command writes.</summary>
*)
{endregion}
METHOD PROTECTED Prepare
VAR
    ObservedState : E_State;
    ObservedExecutionStatus : E_ExecutionStatus;
END_VAR
IF NOT __ISVALIDREF(FResource) THEN
    UpdateStatus(State := E_State.Error,
        ExecutionStatus := E_ExecutionStatus.Error,
        Ready := FALSE);
    RETURN;
END_IF;

IF FResource.HasError THEN
    UpdateStatus(State := E_State.Error,
        ExecutionStatus := E_ExecutionStatus.Error,
        Ready := FALSE);
    RETURN;
END_IF;

IF Enabled AND FResource.IsReady AND (FResource.RequestedValue <> TargetValue) THEN
    FResource.RequestValue(Value := TargetValue);
END_IF;

IF (FResource.ActualValue = TargetValue) AND (FResource.RequestedValue = TargetValue) THEN
    ObservedState := E_State.Completed;
    ObservedExecutionStatus := E_ExecutionStatus.Completed;
ELSIF Enabled AND FResource.IsReady THEN
    ObservedState := E_State.Running;
    ObservedExecutionStatus := E_ExecutionStatus.Running;
ELSIF FResource.IsReady THEN
    ObservedState := E_State.Idle;
    ObservedExecutionStatus := E_ExecutionStatus.Idle;
ELSE
    ObservedState := E_State.Idle;
    ObservedExecutionStatus := E_ExecutionStatus.NotReady;
END_IF;

UpdateStatus(State := ObservedState,
    ExecutionStatus := ObservedExecutionStatus,
    Ready := FResource.IsReady);
END_METHOD

END_FUNCTION_BLOCK

